(* IEC 61131-3 sources: brOscatLib/oscatBasic, 546 files *)

(* ---- oscatBasic.typ ---- *)
TYPE
    REAL2 :    STRUCT
        R1 : REAL; (* small value *)
        RX : REAL; (* big value *)
    END_STRUCT;
    CONSTANTS_LANGUAGE :    STRUCT
        DEFAULT : INT := 1; (* 1=english, 2=german 3=french *)
        LMAX : INT := 3;
        WEEKDAYS : ARRAY[1..3, 1..7] OF STRING[10] := ['Monday', 'Tuesday', 'Wednesday', 'Thursday', 'Friday', 'Saturday', 'Sunday', 'Montag', 'Dienstag', 'Mittwoch', 'Donnerstag', 'Freitag', 'Samstag', 'Sonntag', 'Lundi', 'Mardi', 'Mercredi', 'Jeudi', 'Vendredi', 'Samedi', 'Dimanche'];
        WEEKDAYS2 : ARRAY[1..3, 1..7] OF STRING[2] := ['Mo', 'Tu', 'We', 'Th', 'Fr', 'Sa', 'Su', 'Mo', 'Di', 'Mi', 'Do', 'Fr', 'Sa', 'So', 'Lu', 'Ma', 'Me', 'Je', 'Ve', 'Sa', 'Di'];
        MONTHS : ARRAY[1..3, 1..12] OF STRING[10] := ['January', 'February', 'March', 'April', 'May', 'June', 'July', 'August', 'September', 'October', 'November', 'December', 'Januar', 'Februar', 'März', 'April', 'Mai', 'Juni', 'Juli', 'August', 'September', 'Oktober', 'November', 'Dezember', 'Janvier', 'Février', 'mars', 'Avril', 'Mai', 'Juin', 'Juillet', 'Août', 'Septembre', 'Octobre', 'Novembre', 'Decembre'];
        MONTHS3 : ARRAY[1..3, 1..12] OF STRING[3] := ['Jan', 'Feb', 'Mar', 'Apr', 'May', 'Jun', 'Jul', 'Aug', 'Sep', 'Oct', 'Nov', 'Dec', 'Jan', 'Feb', 'Mrz', 'Apr', 'Mai', 'Jun', 'Jul', 'Aug', 'Sep', 'Okt', 'Nov', 'Dez', 'Jan', 'Fev', 'Mar', 'Avr', 'Mai', 'Jun', 'Jul', 'Aou', 'Sep', 'Oct', 'Nov', 'Dec'];
        DIRS : ARRAY[1..3, 0..15] OF STRING[3] := ['N', 'NNE', 'NE', 'ENE', 'E', 'ESE', 'SE', 'SSE', 'S', 'SSW', 'SW', 'WSW', 'W', 'WNW', 'NW', 'NNW', 'N', 'NNO', 'NO', 'ONO', 'O', 'OSO', 'SO', 'SSO', 'S', 'SSW', 'SW', 'WSW', 'W', 'WNW', 'NW', 'NNW', 'N', 'NNO', 'NO', 'ONO', 'O', 'OSO', 'SO', 'SSO', 'S', 'SSW', 'SW', 'WSW', 'W', 'WNW', 'NW', 'NNW'];
    END_STRUCT;
    CONSTANTS_LOCATION :    STRUCT
        DEFAULT : INT := 1; (* 1=germany, 2=austria 3=france 4=belgium-german 5= italien-Südtirol *)
        LMAX : INT := 5;
        LANGUAGE : ARRAY[1..5] OF INT := [2, 2, 3, 2, 2]; (* language spoken in the location *)
    END_STRUCT;
    CONSTANTS_MATH :    STRUCT
        PI : REAL := 3.1415926535897931; (* Kreiszahl PI *)
        PI2 : REAL := 6.2831853071795862; (* PI * 2 *)
        PI4 : REAL := 12.566370614359172; (* PI * 4 *)
        PI05 : REAL := 1.5707963267949; (* PI / 2 *)
        PI025 : REAL := 0.785398163397448; (* PI / 4 *)
        PI_INV : REAL := 0.318309886183791; (* 1 / PI *)
        E : REAL := 2.7182818284590451; (* Euler constant e *)
        E_INV : REAL := 0.367879441171442; (* 1 / e *)
        SQ2 : REAL := 1.4142135623731; (* Wurzel von 2 *)
        FACTS : ARRAY[0..12] OF DINT := [1, 1, 2, 6, 24, 120, 720, 5040, 40320, 362880, 3628800, 39916800, 479001600];
    END_STRUCT;
    CONSTANTS_PHYS :    STRUCT
        C : REAL := 299792458; (* Lichtgeschwindigkeit in m/s *)
        E : REAL := 1.60217653E-19; (* elementarladung in Colomb = A * s *)
        G : REAL := 9.80665; (* Erdbeschleunigung in m / s² *)
        T0 : REAL := -273.15; (* absoluter Nullpunkt in °C *)
        RU : REAL := 8.314472; (* Universelle Gaskonstante in J / (mol · K) *)
        PN : REAL := 101325; (* NormalDruck in Pa *)
    END_STRUCT;
    CONSTANTS_SETUP :    STRUCT
        EXTENDED_ASCII : BOOL := TRUE; (* setup Parameters *)
        CHARNAMES : ARRAY[1..4] OF STRING[253] := [';"&quot;&&amp;<&lt;>&gt;€&euro; &nbsp;¡&iexcl;¢&cent;£&pound;¤&curren;¥&yen;¦&brvbar;§&sect;¨&uml;©&copy;ª&ordf;«&laquo;¬&not;­&shy;®&reg;¯&macr;°&deg;±&plusmn;²&sup2;³&sup3;´&acute;µ&micro;¶&para;·&middot;¸&cedil;¹&sup1;º&ordm;»&raquo;¼&frac14;Û&Ucirc;',
		';¾&frac34;¿&iquest;À&Agrave;Á&Aacute;Â&Acirc;Ã&Atilde;Ä&Auml;Å&Aring;Æ&AElig;Ç&Ccedil;È&Egrave;É&Eacute;Ê&Ecirc;Ë&Euml;Ì&Igrave;Í&Iacute;Î&Icirc;Ï&Iuml;Ð&ETH;Ñ&Ntilde;Ò&Ograve;Ó&Oacute;Ô&Ocirc;Õ&Otilde;Ö&Ouml;×&times;Ø&Oslash;Ù&Ugrave;Ú&Uacute;½&frac12;',
		';Ü&Uuml;Ý&Yacute;Þ&THORN;ß&szlig;à&agrave;á&aacute;â&acirc;ã&atilde;ä&auml;å&aring;æ&aelig;ç&ccedil;è&egrave;é&eacute;ê&ecirc;ë&euml;ì&igrave;í&iacute;î&icirc;ï&iuml;ð&eth;ñ&ntilde;ò&ograve;ó&oacute;ô&ocirc;õ&otilde;ö&ouml;÷&divide;ø&oslash;ù&ugrave;',
		';ú&uacute;û&ucirc;ü&uuml;ý&yacute;þ&thorn;ÿ&yuml;'];
        MTH_OFS : ARRAY[1..12] OF INT := [0, 31, 59, 90, 120, 151, 181, 212, 243, 273, 304, 334];
        DECADES : ARRAY[0..8] OF REAL := [1, 10, 100, 1000, 10000, 100000, 1000000, 10000000, 100000000];
    END_STRUCT;
    TIMER_EVENT :    STRUCT
        TYP : BYTE;
        CHANNEL : BYTE;
        DAY : BYTE;
        START : TOD;
        DURATION : TIME;
        LAND : BYTE;
        LOR : BYTE;
        LAST : DT;
    END_STRUCT;
    FRACTION :    STRUCT
        NUMERATOR : INT;
        DENOMINATOR : INT;
    END_STRUCT;
    COMPLEX :    STRUCT
        re : REAL;
        im : REAL;
    END_STRUCT;
    VECTOR_3 :    STRUCT
        X : REAL;
        Y : REAL;
        Z : REAL;
    END_STRUCT;
    ESR_DATA :    STRUCT
        TYP : BYTE;
        ADRESS : STRING[10];
        DS : DT;
        TS : TIME;
        DATA : ARRAY[0..7] OF BYTE;
    END_STRUCT;
    CALENDAR :    STRUCT
        UTC : DT; (* world time UTC *)
        LOCAL_DT : DT; (* local time *)
        LOCAL_DATE : DATE; (* local date *)
        LOCAL_TOD : TOD; (* local time of day *)
        YEAR : INT; (* year of LDATE *)
        MONTH : INT; (* month of LDATE *)
        DAY : INT; (* day of LDATE *)
        WEEKDAY : INT; (* weekday of LDATE *)
        OFFSET : INT; (* Time Zone Offset for Local time in minutes *)
        DST_EN : BOOL; (* daylight savings time enable *)
        DST_ON : BOOL; (* true when daylight savings time os on *)
        NAME : STRING[5]; (* name of time zone *)
        LANGUAGE : INT; (* location number pls see location setup *)
        LONGITUDE : REAL; (* longitude of current location *)
        LATITUDE : REAL; (* latitude of current location *)
        SUN_RISE : TOD; (* sun_rise for current location *)
        SUN_SET : TOD; (* sun_set for current location *)
        SUN_MIDDAY : TOD; (* worldtime when sun stands at south position *)
        SUN_HEIGTH : REAL; (* suns heigth at midday, south position *)
        SUN_HOR : REAL; (* sun angle horizontal 0 = north in degrees *)
        SUN_VER : REAL; (* sun angle vertical above horizon in degrees *)
        NIGHT : BOOL; (* true between sun_set and sun_rise *)
        HOLIDAY : BOOL; (* true when holiday *)
        HOLY_NAME : STRING[30]; (* name of holiday *)
        WORK_WEEK : INT; (* current work week *)
    END_STRUCT;
    HOLIDAY_DATA :    STRUCT
        NAME : STRING[30];
        DAY : SINT;
        MONTH : SINT;
        USE : SINT;
    END_STRUCT;
    SDT :    STRUCT
        YEAR : INT;
        MONTH : INT;
        DAY : INT;
        WEEKDAY : INT;
        HOUR : INT;
        MINUTE : INT;
        SECOND : INT;
        MS : INT;
    END_STRUCT;
END_TYPE

(* ---- _ARRAY_ABS.st ---- *)
FUNCTION _ARRAY_ABS
    (*http://www.oscat.de/images/OSCATBasic/oscat_basic333_en.pdf#page=71*)
    stop := SHR(SIZE,2)-1;
    FOR i := 0 TO stop DO
    	PT[i] := ABS(PT[i]);
    END_FOR
    _ARRAY_ABS := TRUE;

    (* revision history
    hm	2. apr 2008		rev 1.0
    	original version

    *)
END_FUNCTION

(* ---- _ARRAY_ADD.st ---- *)
FUNCTION _ARRAY_ADD
    (*http://www.oscat.de/images/OSCATBasic/oscat_basic333_en.pdf#page=71*)
    stop := SHR(SIZE,2)-1;
    FOR i := 0 TO stop DO
    	PT[i] := PT[i] + X;
    END_FOR
    _ARRAY_ADD := TRUE;

    (* revision history
    hm	2. apr 2008		rev 1.0
    	original version

    *)
END_FUNCTION

(* ---- _ARRAY_INIT.st ---- *)
FUNCTION _ARRAY_INIT
    (*http://www.oscat.de/images/OSCATBasic/oscat_basic333_en.pdf#page=72*)
    stop := SHR(SIZE,2)-1;
    FOR i := 0 TO stop DO
    	PT[i] := INIT;
    END_FOR

    _ARRAY_INIT := TRUE;

    (* revision History

    hm 6.1.2007		rev 1.1
    	change type of function to bool
    	added  array_init := true to set output true.

    hm	14.11.2007	rev 1.2
    	changed stop calculation to be more efficient

    hm	16.3. 2008		rev 1.3
    	changed type of input SIZE to uint
    *)
END_FUNCTION

(* ---- _ARRAY_MEDIAN.st ---- *)
FUNCTION _ARRAY_MEDIAN
    (*http://www.oscat.de/images/OSCATBasic/oscat_basic333_en.pdf#page=73*)
    _ARRAY_SORT(ADR(PT),SIZE);
    stop := SHR(SIZE,2)-1;
    IF EVEN(UINT_TO_INT(stop)) THEN
    	_ARRAY_MEDIAN := PT[SHR(stop,1)];
    ELSE
    	i := SHR(stop,1);
    	_ARRAY_MEDIAN := (PT[i] + PT[i+1]) * 0.5;
    END_IF

    (* old code
    stop := (SIZE - SIZEOF(PT)) / SIZEOF(PT);
    FOR i := 0 TO stop - 1 DO
    	FOR m := i + 1 TO stop DO
    		IF PT[i] > PT[m] THEN
    			temp := PT[i];
    			PT[i] := PT[m];
    			PT[m] := temp;
    		END_IF
    	END_FOR
    END_FOR
    IF even(stop) THEN
    	_ARRAY_MEDIAN := PT[stop/2];
    ELSE
    	i := stop/2;
    	_ARRAY_MEDIAN := (PT[i] + PT[i+1])/2;
    END_IF
    *)
    (* revision history
    hm 	3.3.2007		rev 1.1
    	corrected an error, changed the statement line 14	i := TRUNC(stop/2); to i := stop/2;

    hm		22. sep 2007	rev 1.2
    	changed algorithm to use _array_soft for performance reasons

    hm		8. oct 2007		rev 1.3
    	deleted unused variables m and temp

    hm		14. nov 2007	rev 1.4
    	corrected a problem with SIZE calculation

    hm		16.3. 2008		rev 1.5
    	changed type of input SIZE to uint
    	performance improvements
    *)
END_FUNCTION

(* ---- _ARRAY_MUL.st ---- *)
FUNCTION _ARRAY_MUL
    (*http://www.oscat.de/images/OSCATBasic/oscat_basic333_en.pdf#page=73*)
    stop := SHR(SIZE,2)-1;
    FOR i := 0 TO stop DO
    	PT[i] := PT[i] * X;
    END_FOR
    _ARRAY_MUL := TRUE;

    (* revision history
    hm	2. apr 2008		rev 1.0
    	original version

    *)
END_FUNCTION

(* ---- _ARRAY_SHUFFLE.st ---- *)
FUNCTION _ARRAY_SHUFFLE
    (*http://www.oscat.de/images/OSCATBasic/oscat_basic333_en.pdf#page=74*)
    stop := UINT_TO_INT(SHR(SIZE,2)-1);
    FOR i := 0 TO stop DO
            pos := RDM2(i+pos,0,stop);
            (* swap elements *)
            temp := PT[i];
            PT[i] := PT[pos];
            PT[pos] := temp;
    END_FOR

    _ARRAY_SHUFFLE := TRUE;

    (* revision History
    hm 	4. mar 2008	rev 1.0
    	original version

    hm	16. mar. 2008	rev 1.1
    	changed type of input SIZE to uint

    hm	30. mar. 2008	rev 1.2
    	changed last in rdm2 fromm pos to i + pos to allow for more randomness

    *)
END_FUNCTION

(* ---- _ARRAY_SORT.st ---- *)
FUNCTION _ARRAY_SORT
    (*http://www.oscat.de/images/OSCATBasic/oscat_basic333_en.pdf#page=75*)
    (* Startwerte zur Arraygröße *)
    links := 1;					(* Anfangselement des Arrays *)
    rechts := SHR(SIZE,2);		(* Endelement des Arrays *)
    stack_count := 1;			(* Laufvariable stack *)

    WHILE NOT ende_aussen DO						(* äußere Schleife *)
    	IF links < rechts THEN
    		pivot := PT[SHR(rechts+links,1)];			(* Wert des mittleren Elements als pivot-Wert *)
    		i := links -1;
    		j := rechts +1;

    		(* innere Schleife, teile Feld *)
    		ende_innen := FALSE;
    		REPEAT

    			(* steigende Reihenfolge *)
    			REPEAT	i := i+1;	UNTIL (PT[i] >= pivot) OR NOT (i < rechts)	END_REPEAT
    			REPEAT	j := j-1;	UNTIL (PT[j] <= pivot) OR NOT (j > links)	END_REPEAT

    			(*sinkende Reihenfolge *)
    (*			REPEAT	i := i+1;	UNTIL (PT[i] <= pivot) OR NOT (i < rechts)	END_REPEAT	*)
    (*			REPEAT	j := j-1;	UNTIL (PT[j] >= pivot) OR NOT (j > links)	END_REPEAT	*)

    			IF i >= j THEN
    				ende_innen := TRUE;
    			ELSE
    				   tmp := PT[j];
    				PT[j] := PT[i];
    				PT[i] := tmp;
    			END_IF

    		UNTIL ende_innen END_REPEAT

    		(* Push stack *)
    		stack[stack_count] := rechts;		(* rechten Teil später sortieren *)
    		IF stack_count < 32 THEN
    			stack_count := stack_count +1;
    		ELSE
    			ende_aussen := TRUE;
    			_ARRAY_SORT := FALSE;					(* Fehler: stack zu klein *)
    		END_IF

    		(* linken Teil sortiern *)
    		rechts := MAX(links, i-1);

    	ELSE

    		IF stack_count = 1 THEN
    			ende_aussen := TRUE;
    		ELSE

    			links := rechts+1;

    			(* pop stack *)
    			stack_count := stack_count -1;		(* jetzt rechten Teil sortierne *)
    			rechts:= stack[stack_count];
    		END_IF

    	END_IF

    END_WHILE

    _ARRAY_SORT := TRUE;				(* Sortierung beendet *)

    (* algorithm used before rev 2.0

    SIZE := SHR(SIZE,2);
    size2 := UINT_TO_INT(SHR(SIZE,1));
    FOR i := SIZE2  TO 1 BY -1 DO
    	j:=i;
        WHILE j <= SIZE2 DO
         	stop := j * 2 + 1;
            IF stop > UINT_TO_INT(SIZE) THEN stop := stop - 1;
            ELSIF PT[stop-1] > PT[stop] THEN stop := stop - 1;
    		END_IF
            IF PT[j] < PT[stop] THEN
             	temp := PT[j];
                PT[j] := PT[stop];
                PT[stop] := temp;
            END_IF
            j := stop;
        END_WHILE
    END_FOR

    *)

    (* heapsort
    FOR heapsize := UINT_TO_INT(SIZE) TO 1 BY -1 DO
    	popmax := PT[1];
    	PT[1] := PT[heapsize];
       	i := 1;
    	hs2 := SHR(heapsize,1);
    	WHILE i <= hs2 DO
           	stop := i * 2 + 1;
            	IF stop > heapsize THEN stop := stop - 1;
            	ELSIF PT[stop-1] > PT[stop] THEN stop := stop - 1;
    	 	END_IF
            	IF PT[i] < PT[stop] THEN
                		temp := PT[i];
                		PT[i] := PT[stop];
                		PT[stop] := temp;
            	END_IF
            	i := stop;
        	END_WHILE
    	PT[heapsize] := popmax;
    END_FOR

    _ARRAY_SORT2 := TRUE;
    *)

    (* old algorithm bubble sort used before rev 1.2
    stop := (SIZE - SIZEOF(PT)) / SIZEOF(PT);
    FOR i := 0 TO stop - 1 DO
    	FOR m := i + 1 TO stop DO
    		IF PT[i] > PT[m] THEN
    			temp := PT[i];
    			PT[i] := PT[m];
    			PT[m] := temp;
    		END_IF
    	END_FOR
    END_FOR
    _ARRAY_SORT := TRUE;

    *)

    (* revision history

    hm 	6.1.2007 	rev 1.1
    	changed return value to true

    hm	22. sep 2007	rev 1.2
    	changed sorting algorithm to heap sort for performance reasons

    hm 	14. nov 2007	rev 1.3
    	changed calculation of stop to be more efficient

    hm	15 dec 2007	rev 1.4
    	added function return true

    hm	5. jan 2008		rev 1.5
    	improved performance

    hm	16. mar. 2008	rev 1.6
    	changed type of input SIZE to uint

    hm	28. mar. 2008	rev 1.7
    	changed input f to PT

    hm	19. jan. 2011	rev 2.0
    	new faster algorithm using qucksort (Alexander Drikitis)

    *)

END_FUNCTION

(* ---- _BUFFER_CLEAR.st ---- *)
FUNCTION _BUFFER_CLEAR
    (*http://www.oscat.de/images/OSCATBasic/oscat_basic333_en.pdf#page=477*)
    (* this routine uses 32 bit access to gain speed *)
    (* first access bytes till pointer is aligned for 32 bit access *)
    temp := ADR(PT);
    end := temp + SIZE;
    end32 := end - 3;
    WHILE (ADR(PT) < end) AND ((temp AND 16#00000003) > 0) DO
    	PT := 0;
    	PT ACCESS (ADR(PT) + 1);
    	temp := temp + 1;
    END_WHILE
    (* pointer is aligned, now copy 32 bits at a time *)
    ptw ACCESS ADR(PT);
    WHILE ADR(ptw) < end32 DO (* *)
    	ptw := 0;
    	ptw ACCESS (ADR(ptw) + 4);
    END_WHILE
    (* copy the remaining bytes in byte mode *)
    PT ACCESS ADR(ptw);
    WHILE ADR(PT) < end DO
    	PT := 0;
    	PT ACCESS (ADR(PT) + 1);
    END_WHILE

    _BUFFER_CLEAR := TRUE;

    (* revision History
    hm 	5. mar. 2008	rev 1.0
    	original version

    hm	16. mar. 2008	rev 1.1
    	added type conversion to avoid warnings under codesys 30
    	chaged type of input SIZE to uint
    	deleted unused variable i

    hm	31. oct. 2008	rev 1.2
    	corrected an error while routine would write outside of arrays

    *)
END_FUNCTION

(* ---- _BUFFER_INIT.st ---- *)
FUNCTION _BUFFER_INIT
    (*http://www.oscat.de/images/OSCATBasic/oscat_basic333_en.pdf#page=477*)
    (* this routine uses 32 bit access to gain speed *)
    (* first access bytes till pointer is aligned for 32 bit access *)
    temp := ADR(PT);
    end := temp + SIZE;
    end32 := end - 3;
    WHILE (ADR(PT) < end) AND ((temp AND 16#00000003) > 0) DO
    	PT := INIT;
        PT ACCESS (ADR(PT) + 1);
    	temp := temp + 1;
    END_WHILE
    (* pointer is aligned, now copy 32 bits at a time *)
    ptw ACCESS ADR(PT);
    temp := SHL(BYTE_TO_UDINT(INIT),24) OR SHL(BYTE_TO_UDINT(INIT),16) OR SHL(BYTE_TO_UDINT(INIT),8) OR BYTE_TO_UDINT(INIT);
    WHILE ADR(ptw) < end32 DO
    	ptw := UDINT_TO_DWORD(temp);
    	ptw ACCESS (ADR(ptw) + 4);
    END_WHILE
    (* copy the remaining bytes in byte mode *)
    PT ACCESS ADR(ptw);
    WHILE ADR(PT) < end DO
    	PT := INIT;
    	PT ACCESS (ADR(PT) + 1);
    END_WHILE

    _BUFFER_INIT := TRUE;

    (* revision History
    hm 	5. mar. 2008	rev 1.0
    	original version

    hm	16. mar. 2008	rev 1.1
    	added type conversion to avoid warnings under codesys 3.0
    	chaged type of input SIZE to uint.

    hm	31. oct. 2008	rev 1.2
    	corrected an error while routine would write outside of arrays

    *)
END_FUNCTION

(* ---- _BUFFER_INSERT.st ---- *)
FUNCTION _BUFFER_INSERT
    (*http://www.oscat.de/images/OSCATBasic/oscat_basic333_en.pdf#page=478*)
    lx := LEN(STR);
    end := POS + lx;
    (* first move the upper part of the buffer to make space for the string *)
    FOR i := UINT_TO_INT(SIZE) - 1 TO end BY -1 DO
    	PT[i] := PT[i-lx];
    END_FOR
    (* copy the string *)
    _BUFFER_INSERT := _STRING_TO_BUFFER(STR, POS, ADR(PT), SIZE);

    (* revision History
    hm 	9. mar. 2008	rev 1.0
    	original version

    hm	16. mar. 2008	rev 1.1
    	changed type of input SIZE to uint

    hm	13. may. 2008	rev 1.2
    	changed type of pointer to array[1..32767]
    	changed SIZE of string to STRING_LENGTH

    hm	23. mar. 2009	rev 1.3
    	avoid writing to input POS

    hm	12. nov. 2009	rev 1.4
    	code optimized

    hm 2. jan 2012	rev 1.5
    	function now returns the next position after the input string

    *)
END_FUNCTION

(* ---- _BUFFER_UPPERCASE.st ---- *)
FUNCTION _BUFFER_UPPERCASE
    (*http://www.oscat.de/images/OSCATBasic/oscat_basic333_en.pdf#page=479*)
    pos := 0;
    WHILE pos < SIZE DO
    	PT[pos] := TO_UPPER(PT[pos]);
    	pos := pos + 1;
    END_WHILE

    _BUFFER_UPPERCASE := TRUE;

    (* revision History
    hm 	20. jan. 2011	rev 1.0
    	original version

    *)
END_FUNCTION

(* ---- _STRING_TO_BUFFER.st ---- *)
FUNCTION _STRING_TO_BUFFER
    (*http://www.oscat.de/images/OSCATBasic/oscat_basic333_en.pdf#page=479*)
    ps ACCESS ADR(STR);
    end := MIN(POS + LEN(STR), UINT_TO_INT(SIZE));
    IF end > 0 THEN end := end -1; END_IF
    FOR i := POS TO end DO
    	PT[i] := ps;
    	ps ACCESS (ADR(ps) + 1);
    END_FOR

    _STRING_TO_BUFFER := i;

    (* revision History

    hm 	5. mar. 2008	rev 1.0
    	original version

    hm	16. mar. 2008	rev 1.1
    	changed type of input SIZE to uint

    hm	13. may. 2008	rev 1.2
    	changed type of pointer to array[1..32767]
    	changed SIZE of string to STRING_LENGTH

    hm	12. nov. 2009	rev 1.3
    	limit end to SIZE - 1

    hm	2. jan 2012	rev 1.4
    	return the position after the input string when finished
    *)
END_FUNCTION

(* ---- ACOSH.st ---- *)
FUNCTION ACOSH
    (*http://www.oscat.de/images/OSCATBasic/oscat_basic333_en.pdf#page=39*)
    ACOSH := LN(SQRT(X * X - 1.0) + X);

    (* revision history
    hm		12 jan 2007	rev 1.0
    	original version

    hm		2. dec 2007	rev 1.1
    	changed code for better performance

    hm	16. mar. 2007		rev 1.2
    	changed sequence of calculations to improve performance

    hm	10. mar. 2009		rev 1.3
    	real constants updated to new systax using dot

    *)
END_FUNCTION

(* ---- ACOTH.st ---- *)
FUNCTION ACOTH
    (*http://www.oscat.de/images/OSCATBasic/oscat_basic333_en.pdf#page=39*)
    ACOTH := LN((X+1.0)/(X-1.0))*0.5;

    (* revision history
    hm		12 jan 2007	rev 1.0
    	original version

    hm		5. jan 2008	rev 1.1
    	improved code for better performance

    hm	10. mar. 2009		rev 1.2
    	real constants updated to new systax using dot

    *)
END_FUNCTION

(* ---- AGDF.st ---- *)
FUNCTION AGDF
    (*http://www.oscat.de/images/OSCATBasic/oscat_basic333_en.pdf#page=39*)
    AGDF := LN((1.0 + SIN(X)) / COS(X));

    (* comment
    the current implementation gives sufficient accuracy only up to X = 1.57 or an output > 10.
    is X closer to PI/2 then the function is more and more unreliable
    *)

    (* revision history
    hm	27. apr. 2008	rev 1.0
    	original version

    hm	10. mar. 2009	rev 1.1
    	real constants updated to new systax using dot

    *)

END_FUNCTION

(* ---- AIN.st ---- *)
FUNCTION AIN
    (*http://www.oscat.de/images/OSCATBasic/oscat_basic333_en.pdf#page=269*)
    (* extract the SIGN bit *)
    IF SIGN < 32 THEN
    	temp1 := SHR(IN,SIGN);
    	sx := temp1.0;
    ELSE
    	sx := FALSE;
    END_IF
    temp1 := SHR(ff, 32-BYTE_TO_USINT(BITS));
    temp2 := IN AND temp1;
    AIN := (HIGH - LOW) * DWORD_TO_REAL(temp2) / DWORD_TO_REAL(temp1) + LOW;
    IF sx THEN AIN := -AIN; END_IF

    (* revision history
    hm 18.8.2006	rev 1.1
    	fixed an error with LOW value negative and HIGH value 0.

    hm 19.1.2007	rev 1.2
    	fixed an error with SIGN bit.

    hm	13.9.2007	rev 1.3
    	changed code to avoid warning under codesys 2.8.1

    hm	2. dec 2007	rev 1.4
    	changed code for better performance

    hm	16. mar 2008	rev 1.5
    	added type conversions to avoid warnings under codesys 30
    *)
END_FUNCTION

(* ---- AOUT.st ---- *)
FUNCTION AOUT
    (*http://www.oscat.de/images/OSCATBasic/oscat_basic333_en.pdf#page=271*)
    (* if SIGN bit is defined *)
    IF SIGN < 32 THEN
    	sx := SIGN_R(IN);
    	in2 := ABS(IN);
    ELSE
    	in2 := IN;
    END_IF

    (* begrenze IN auf die zulässigen werte *)
    in2 := LIMIT(LOW, in2, HIGH);

    (* Berechne den Ausgangswert *)
    AOUT := REAL_TO_DWORD((in2 - LOW) / (HIGH - LOW) * UDINT_TO_REAL(SHL(ff,BYTE_TO_USINT(BITS)) -1));
    IF sx THEN AOUT := UDINT_TO_DWORD(SHL(ff,SIGN) OR DWORD_TO_UDINT(AOUT)); END_IF

    (*
    revision history

    hm 18.1.2007		rev 1.1
    	renamed Modul to AOUT.
    	changed Output to 32 Bit max.
    	corrected error with SIGN bit.

    hm	13.9.2007		rev 1.2
    	changed code to avoid warning under codesys 2.8.1

    hm	2. dec 2007		rev 1.3
    	changed code for better performance

    hm	23. feb 2008	rev 1.4
    	changed code for better performance
    *)
END_FUNCTION

(* ---- AOUT1.st ---- *)
FUNCTION AOUT1
    (*http://www.oscat.de/images/OSCATBasic/oscat_basic333_en.pdf#page=272*)
    (* if SIGN bit is defined *)
    IF SIGN < 32 THEN
    	sx := SIGN_R(IN);
    	in2 := ABS(IN);
    ELSE
    	in2 := IN;
    END_IF

    (* begrenze IN auf die zulässigen werte *)
    in2 := LIMIT(LOW, in2, HIGH);

    (* Berechne den Ausgangswert *)
    AOUT1 := SHL(REAL_TO_DWORD((in2 - LOW) / (HIGH - LOW) * UDINT_TO_REAL(SHL(ff,BIT_N - BIT_0 + 1) -1)),BIT_0);
    IF sx THEN AOUT1 := UDINT_TO_DWORD(SHL(ff,SIGN) OR DWORD_TO_UDINT(AOUT1)); END_IF

    (* revision history
    hm	23. feb 2008	rev 1.0
    	original version

    *)
END_FUNCTION

(* ---- ARRAY_AVG.st ---- *)
FUNCTION ARRAY_AVG
    (*http://www.oscat.de/images/OSCATBasic/oscat_basic333_en.pdf#page=76*)
    stop := SHR(SIZE,2)-1;
    ARRAY_AVG := PT[0];
    FOR i := 1 TO stop DO
    	ARRAY_AVG := ARRAY_AVG + PT[i];
    END_FOR
    ARRAY_AVG := ARRAY_AVG / UINT_TO_REAL(stop + 1);

    (* revision history
    hm	2. oct 2007		rev 1.0
    	original version

    hm	12. dec 2007	rev 1.1
    	chaged code for better performance

    hm	16. mar. 2008	rev 1.2
    	changed input SIZE to uint

    hm	10. mar. 2009	rev 1.3
    	added type conversion for compatibility reasons
    *)
END_FUNCTION

(* ---- ARRAY_GAV.st ---- *)
FUNCTION ARRAY_GAV
    (*http://www.oscat.de/images/OSCATBasic/oscat_basic333_en.pdf#page=76*)
    stop := SHR(SIZE,2)-1;
    ARRAY_GAV := 1.0;
    FOR i := 0 TO stop DO
    	IF PT[i] > 0.0 THEN
    		ARRAY_GAV := ARRAY_GAV * PT[i];
    	ELSE
    		ARRAY_GAV := 0.0;
    		RETURN;
    	END_IF
    END_FOR
    ARRAY_GAV := SQRTN(ARRAY_GAV,UINT_TO_INT(stop)+1);

    (* revision history
    hm	2. apr 2008	rev 1.0
    	original version

    hm	10. mar. 2009	rev 1.1
    	real constants updated to new systax using dot

    *)
END_FUNCTION

(* ---- ARRAY_HAV.st ---- *)
FUNCTION ARRAY_HAV
    (*http://www.oscat.de/images/OSCATBasic/oscat_basic333_en.pdf#page=77*)
    stop := SHR(SIZE,2)-1;
    FOR i := 0 TO stop DO
    	IF PT[i] <> 0.0 THEN
    		ARRAY_HAV := ARRAY_HAV + 1.0 / PT[i];
    	ELSE
    		ARRAY_HAV := 0.0;
    		RETURN;
    	END_IF
    END_FOR
    ARRAY_HAV := UINT_TO_REAL(stop + 1) / ARRAY_HAV;

    (* revision history
    hm	2. apr 2008	rev 1.0
    	original version

    hm	10. mar. 2009	rev 1.1
    	real constants updated to new systax using dot

    *)
END_FUNCTION

(* ---- ARRAY_MAX.st ---- *)
FUNCTION ARRAY_MAX
    (*http://www.oscat.de/images/OSCATBasic/oscat_basic333_en.pdf#page=77*)
    stop := (SIZE -SIZEOF(PT)) / SIZEOF(PT);
    ARRAY_MAX := PT[0];
    FOR i := 1 TO stop DO
    	IF PT[i] > ARRAY_MAX THEN ARRAY_MAX := PT[i]; END_IF
    END_FOR

    (* revision history
    hm	2. oct 2006		rev 1.0
    	original version

    hm	16. mar. 2008	rev 1.1
    	changed input SIZE to uint
    *)
END_FUNCTION

(* ---- ARRAY_MIN.st ---- *)
FUNCTION ARRAY_MIN
    (*http://www.oscat.de/images/OSCATBasic/oscat_basic333_en.pdf#page=78*)
    stop := (SIZE - SIZEOF(PT)) / SIZEOF(PT);
    ARRAY_MIN := PT[0];
    FOR i := 1 TO stop DO
    	IF PT[i] < ARRAY_MIN THEN ARRAY_MIN := PT[i]; END_IF
    END_FOR

    (* revision history
    hm		2. oct. 2006
    	original version

    hm		16. mar. 2008
    	changed type of input SIZE to uint

    *)
END_FUNCTION

(* ---- ARRAY_SDV.st ---- *)
FUNCTION ARRAY_SDV
    (*http://www.oscat.de/images/OSCATBasic/oscat_basic333_en.pdf#page=79*)
    (* standard deviation is simply the square root of the variance *)

    ARRAY_SDV := SQRT(ARRAY_VAR(ADR(PT), SIZE));

    (* revision history
    hm 	1.4.2007		rev 1.0
    	function created

    hm	16. mar. 2008	rev 1.1
    	changed type of input SIZE to uint

    *)
END_FUNCTION

(* ---- ARRAY_SPR.st ---- *)
FUNCTION ARRAY_SPR
    (*http://www.oscat.de/images/OSCATBasic/oscat_basic333_en.pdf#page=79*)
    stop := (SIZE -SIZEOF(PT)) / SIZEOF(PT);
    array_min := PT[0];
    array_max := PT[0];
    FOR i := 1 TO stop DO
    	IF PT[i] > array_max THEN array_max := PT[i];
    	ELSIF PT[i] < array_min THEN array_min := PT[i];
    	END_IF
    END_FOR
    ARRAY_SPR := array_max - array_min;

    (* revision history
    hm 	2. oct. 2006	rev 1.0
    	original version

    hm	16. mar. 2008	rev 1.1
    	changed type of input SIZE to uint

    *)
END_FUNCTION

(* ---- ARRAY_SUM.st ---- *)
FUNCTION ARRAY_SUM
    (*http://www.oscat.de/images/OSCATBasic/oscat_basic333_en.pdf#page=80*)
    stop := (SIZE -SIZEOF(PT)) / SIZEOF(PT);
    ARRAY_SUM := PT[0];
    FOR i := 1 TO stop DO
    	ARRAY_SUM := ARRAY_SUM + PT[i];
    END_FOR

    (* revision history
    hm 	2. oct. 2006	rev 1.0
    	function created

    hm	16. mar. 2008	rev 1.1
    	changed type of input SIZE to uint

    *)
END_FUNCTION

(* ---- ARRAY_TREND.st ---- *)
FUNCTION ARRAY_TREND
    (*http://www.oscat.de/images/OSCATBasic/oscat_basic333_en.pdf#page=81*)
    stop := SHR(SIZE,2)-1;
    stop2 := SHR(stop,1);
    FOR i := 0 TO stop2 DO x := x - PT[i]; END_FOR
    IF EVEN(UINT_TO_INT(stop)) THEN
    	FOR i := stop2 TO stop DO x := x + PT[i]; END_FOR
    ELSE
    	FOR i := stop2 + 1 TO stop DO x := x + PT[i]; END_FOR
    END_IF
    ARRAY_TREND := x / UINT_TO_REAL(stop2 + 1);

    (* revision history
    hm	2 oct 2007	rev 1.0
    	original version

    hm	12 dec 2007	rev 1.1
    	changed code for better performance

    hm	16. mar. 2008	rev 1.2
    	changed type of input SIZE to uint

    hm	10. mar. 2009	rev 1.3
    	added type conversions for compatibility reasons
    *)
END_FUNCTION

(* ---- ARRAY_VAR.st ---- *)
FUNCTION ARRAY_VAR
    (*http://www.oscat.de/images/OSCATBasic/oscat_basic333_en.pdf#page=81*)
    (* at first we calualte the arithmetic average of the array *)

    stop := SHR(SIZE,2)-1;
    avg := PT[0];
    FOR i := 1 TO stop DO
    	avg := avg + PT[i];
    END_FOR
    avg := avg / UINT_TO_REAL(stop + 1);

    (* in a second run we calculate the variance of the array *)

    ARRAY_VAR := (PT[0] - avg) * (PT[0] - avg);
    FOR i := 1 TO stop DO
    	ARRAY_VAR := ARRAY_VAR + (PT[i] - avg) * (PT[i] - avg);
    END_FOR
    ARRAY_VAR := ARRAY_VAR / UINT_TO_REAL(stop);

    (* revision history
    hm 	1.4.2007	rev 1.0
    	function created

    hm	12.12.2007	rev 1.1
    	changed code for better performance

    hm	16. mar. 2008	rev 1.2
    	changed type of input SIZE to uint

    hm	10. mar. 2009	rev 1.3
    	added type conversions for compatibility reasons
    *)
END_FUNCTION

(* ---- ASINH.st ---- *)
FUNCTION ASINH
    (*http://www.oscat.de/images/OSCATBasic/oscat_basic333_en.pdf#page=40*)
    ASINH := LN(SQRT(X * X + 1.0)+X);

    (* revision history
    hm		12 jan 2007	rev 1.0
    	original version

    hm		2. dec 2007	rev 1.1
    	changed code for better performance

    hm		16.3. 2007		rev 1.2
    	changed sequence of calculations to improve performance

    hm	10. mar. 2009		rev 1.3
    	real constants updated to new systax using dot

    *)
END_FUNCTION

(* ---- ATAN2.st ---- *)
FUNCTION ATAN2
    (*http://www.oscat.de/images/OSCATBasic/oscat_basic333_en.pdf#page=40*)
    IF X > 0.0 THEN
    	ATAN2 := ATAN(Y/X);
    ELSIF X < 0.0 THEN
    	IF Y >=0.0 THEN
    		ATAN2 := ATAN(Y/X) + cPI;
    	ELSE
    		ATAN2 := ATAN(Y/X) - cPI;
    	END_IF
    ELSIF Y > 0.0 THEN
    	ATAN2 := cPI05;
    ELSIF Y < 0.0 THEN
    	ATAN2 := -cPI05;
    ELSE
    	ATAN2 := 0.0;
    END_IF

    (* revision history
    hm	20.  apr. 2008	rev 1.0
    	original version

    hm	18. oct. 2008	rev 1.1
    	changed to use math constants

    hm	10. mar. 2009	rev 1.2
    	real constants updated to new systax using dot

    *)

END_FUNCTION

(* ---- ATANH.st ---- *)
FUNCTION ATANH
    (*http://www.oscat.de/images/OSCATBasic/oscat_basic333_en.pdf#page=41*)
    ATANH := LN((1.0 + X)/(1.0 - X)) * 0.5;

    (* revision history
    hm		12 jan 2007	rev 1.0
    	original version

    hm		5. jan 2008	rev 1.1
    	improved code for better performance

    hm	10. mar. 2009		rev 1.2
    	real constants updated to new systax using dot

    *)

END_FUNCTION

(* ---- BAND_B.st ---- *)
FUNCTION BAND_B
    (*http://www.oscat.de/images/OSCATBasic/oscat_basic333_en.pdf#page=377*)
    IF BYTE_TO_SINT(X) < BYTE_TO_SINT(B) THEN
    	BAND_B := 0;
    ELSIF BYTE_TO_SINT(X) > (255 - BYTE_TO_SINT(B)) THEN
    	BAND_B := 255;
    ELSE
    	BAND_B := X;
    END_IF

    (* revision history
    hm	21. nov. 2008	rev 1.0
    	original version

    *)

END_FUNCTION

(* ---- BCDC_TO_INT.st ---- *)
FUNCTION BCDC_TO_INT
    (*http://www.oscat.de/images/OSCATBasic/oscat_basic333_en.pdf#page=210*)
    BCDC_TO_INT := (BYTE_TO_INT(IN) AND 16#0F) + (SHR(BYTE_TO_INT(IN),4) * 10);

    (* revision history
    hm	13.12.2007	rev 1.0
    	original version

    hm	30.6.2008	rev 1.1
    	changed name BCD_TO_INT to BCDC_TO_INT to avoid collision with util.lib

    *)
END_FUNCTION

(* ---- BETA.st ---- *)
FUNCTION BETA
    (*http://www.oscat.de/images/OSCATBasic/oscat_basic333_en.pdf#page=41*)
    BETA := GAMMA(X) * GAMMA(Y) / GAMMA(X + Y);

    (* revision history
    hm	26. oct. 2008	rev 1.0
    	original version

    *)
END_FUNCTION

(* ---- BFT_TO_MS.st ---- *)
FUNCTION BFT_TO_MS
    (*http://www.oscat.de/images/OSCATBasic/oscat_basic333_en.pdf#page=354*)
    BFT_TO_MS := EXPT(BFT, 1.5) * 0.836;

    (* revision history
    hm	12. 6. 2008		rev 1.0
    	original version

    *)
END_FUNCTION

(* ---- BIN_TO_BYTE.st ---- *)
FUNCTION BIN_TO_BYTE
    (*http://www.oscat.de/images/OSCATBasic/oscat_basic333_en.pdf#page=145*)
    pt ACCESS ADR(BIN);
    stop := LEN(BIN);
    FOR i := 1 TO stop DO
    	X := pt;
    	(* calculate the value of the digit *)
    	IF X = BYTE#48 THEN
    		BIN_TO_BYTE := SHL(BIN_TO_BYTE,1);
    	ELSIF X = BYTE#49 THEN
    		BIN_TO_BYTE := SHL(BIN_TO_BYTE,1) OR 1;
    	END_IF
    	pt ACCESS (ADR(pt) + 1);
    END_FOR

    (* revision histroy
    hm	18. jun. 2008	rev 1.0
    	original release

    hm	20. sep. 2008	rev 1.1
    	changed length of input string from 20 to 12

    hm	26. jul. 2009	rev 1.2
    	optimized code
    *)

END_FUNCTION

(* ---- BIN_TO_DWORD.st ---- *)
FUNCTION BIN_TO_DWORD
    (*http://www.oscat.de/images/OSCATBasic/oscat_basic333_en.pdf#page=145*)
    pt ACCESS ADR(BIN);
    stop := LEN(BIN);
    FOR i := 1 TO stop DO
    	X := pt;
    	(* calculate the value of the digit *)
    	IF X = BYTE#48 THEN
    		BIN_TO_DWORD := SHL(BIN_TO_DWORD,1);
    	ELSIF X = BYTE#49 THEN
    		BIN_TO_DWORD := SHL(BIN_TO_DWORD,1) OR 1;
    	END_IF
    	pt ACCESS (ADR(pt) + 1);
    END_FOR

    (* revision histroy
    hm	18. jun. 2008	rev 1.0
    	original release

    hm	20. sep. 2008	rev 1.1
    	changed length of input dtring from 20 to 40

    hm	26. jul 2009	rev 1.2
    	optimized code
    *)

END_FUNCTION

(* ---- BINOM.st ---- *)
FUNCTION BINOM
    (*http://www.oscat.de/images/OSCATBasic/oscat_basic333_en.pdf#page=42*)
    IF 2 * K > N THEN
    	K := N - K;
    END_IF
    IF K > N THEN
    	RETURN;
    ELSIF K = 0 OR K = N THEN
    	BINOM := 1;
    ELSIF K = 1 THEN
    	BINOM := N;
    ELSE
    	BINOM := N;
    	N := N + 1;
    	FOR i := 2 TO K DO
    		BINOM := BINOM * (N - i) / i;
    	END_FOR
    END_IF

    (*
    binomialkoeffizient(N, K)
    1  wenn K = 0 return 1
    2  wenn 2k > N
    3      dann führe aus ergebnis \leftarrow binomialkoeffizient(N, N-K)
    4  sonst führe aus ergebnis \leftarrow N
    5          von i \leftarrow 2 bis K
    6              führe aus ergebnis \leftarrow ergebnis \cdot (N + 1 - i)
    7                        ergebnis \leftarrow ergebnis : i
    8  return ergebnis
    *)

    (* revision history
    hm	25. oct. 2008	rev 1.0
    	original version

    *)
END_FUNCTION

(* ---- BIT_COUNT.st ---- *)
FUNCTION BIT_COUNT
    (*http://www.oscat.de/images/OSCATBasic/oscat_basic333_en.pdf#page=210*)
    WHILE IN > 0 DO
    	IF IN.0 THEN BIT_COUNT := BIT_COUNT + 1; END_IF
    	IN := SHR(IN,1);
    END_WHILE

    (* revision history
    5.7.2007	rev 1.0		original version

    10.9.2007	rev 1.1		hm
    	changed algorithm for better performace
    	the execution time has reduced by a factor of 5
    	deleted unused variable temp
    *)
END_FUNCTION

(* ---- BIT_LOAD_B.st ---- *)
FUNCTION BIT_LOAD_B
    (*http://www.oscat.de/images/OSCATBasic/oscat_basic333_en.pdf#page=210*)
    IF VAL THEN
    	BIT_LOAD_B := IN OR SHL(dat,POS);
    ELSE
    	BIT_LOAD_B := IN AND (NOT SHL(dat,POS));
    END_IF

    (* revision history
    hm	29. feb 2008	rev 1.0
    	original version

    hm	16. mar 2008	rev 1.1
    	change input bit to VAL for compatibility reasons
    *)

END_FUNCTION

(* ---- BIT_LOAD_B2.st ---- *)
FUNCTION BIT_LOAD_B2
    (*http://www.oscat.de/images/OSCATBasic/oscat_basic333_en.pdf#page=211*)
    IF D THEN
    	BIT_LOAD_B2 := ROL(SHR(BYTE#255, 8 - N) OR ROR(I, P), P);
    ELSE
    	BIT_LOAD_B2 := ROL(SHL(BYTE#255, N) AND ROR(I, P), P);
    END_IF

    (* revision history
    hm	18. oct. 2008	rev 1.0
    	original version

    *)

END_FUNCTION

(* ---- BIT_LOAD_DW.st ---- *)
FUNCTION BIT_LOAD_DW
    (*http://www.oscat.de/images/OSCATBasic/oscat_basic333_en.pdf#page=211*)
    IF VAL THEN
    	BIT_LOAD_DW := IN OR SHL(dat,POS);
    ELSE
    	BIT_LOAD_DW := IN AND (NOT SHL(dat,POS));
    END_IF

    (* revision history
    hm	29. feb 2008	rev 1.0
    	original version

    hm	16. mar 2008	rev 1.1
    	change input bit to VAL for compatibility reasons
    *)

END_FUNCTION

(* ---- BIT_LOAD_DW2.st ---- *)
FUNCTION BIT_LOAD_DW2
    (*http://www.oscat.de/images/OSCATBasic/oscat_basic333_en.pdf#page=212*)
    IF D THEN
    	BIT_LOAD_DW2 := ROL(SHR(DWORD#4294967295, 32 - N) OR ROR(I, P), P);
    ELSE
    	BIT_LOAD_DW2 := ROL(SHL(DWORD#4294967295, N) AND ROR(I, P), P);
    END_IF

    (* revision history
    hm	18. oct. 2008	rev 1.0
    	original version

    *)

END_FUNCTION

(* ---- BIT_LOAD_W.st ---- *)
FUNCTION BIT_LOAD_W
    (*http://www.oscat.de/images/OSCATBasic/oscat_basic333_en.pdf#page=212*)
    IF VAL THEN
    	BIT_LOAD_W := IN OR SHL(dat,POS);
    ELSE
    	BIT_LOAD_W := IN AND (NOT SHL(dat,POS));
    END_IF

    (* revision history
    hm	29. feb 2008	rev 1.0
    	original version

    hm	16. mar 2008	rev 1.1
    	change input bit to VAL for compatibility reasons
    *)

END_FUNCTION

(* ---- BIT_LOAD_W2.st ---- *)
FUNCTION BIT_LOAD_W2
    (*http://www.oscat.de/images/OSCATBasic/oscat_basic333_en.pdf#page=213*)
    IF D THEN
    	BIT_LOAD_W2 := ROL(SHR(WORD#65535, 16 - N) OR ROR(I, P), P);
    ELSE
    	BIT_LOAD_W2 := ROL(SHL(WORD#65535, N) AND ROR(I, P), P);
    END_IF

    (* revision history
    hm	18. oct. 2008	rev 1.0
    	original version

    *)

END_FUNCTION

(* ---- BIT_OF_DWORD.st ---- *)
FUNCTION BIT_OF_DWORD
    (*http://www.oscat.de/images/OSCATBasic/oscat_basic333_en.pdf#page=213*)
    BIT_OF_DWORD := (SHR(IN,N) AND 16#00000001) > 0;

    (* old code used before rev 1.1
    temp := SHR(IN,N);
    BIT_OF_DWORD := temp.0;
    *)

    (* revision history
    hm	4. aug. 2006	rev 1.0
    	original version

    hm	29. feb 2008	rev 1.1
    	improved performance

    hm	6. jun. 2008	rev 1.2
    	changes type of input N from byte to int
    *)

END_FUNCTION

(* ---- BIT_TOGGLE_B.st ---- *)
FUNCTION BIT_TOGGLE_B
    (*http://www.oscat.de/images/OSCATBasic/oscat_basic333_en.pdf#page=214*)
    BIT_TOGGLE_B := SHL(BYTE#1, POS) XOR IN;

    (* revision history
    hm	18. oct. 2008	rev 1.0
    	original version

    *)

END_FUNCTION

(* ---- BIT_TOGGLE_DW.st ---- *)
FUNCTION BIT_TOGGLE_DW
    (*http://www.oscat.de/images/OSCATBasic/oscat_basic333_en.pdf#page=214*)
    BIT_TOGGLE_DW := SHL(DWORD#1, POS) XOR IN;

    (* revision history
    hm	18. oct. 2008	rev 1.0
    	original version

    *)

END_FUNCTION

(* ---- BIT_TOGGLE_W.st ---- *)
FUNCTION BIT_TOGGLE_W
    (*http://www.oscat.de/images/OSCATBasic/oscat_basic333_en.pdf#page=215*)
    BIT_TOGGLE_W := SHL(WORD#1, POS) XOR IN;

    (* revision history
    hm	18. oct. 2008	rev 1.0
    	original version

    *)

END_FUNCTION

(* ---- BUFFER_COMP.st ---- *)
FUNCTION BUFFER_COMP
    (*http://www.oscat.de/images/OSCATBasic/oscat_basic333_en.pdf#page=480*)
    (* search for first character match *)
    IF SIZE2 <= SIZE1 THEN
    	end := SIZE1 - SIZE2;
    	firstbyte := PT2[0];
    	FOR i := START TO end DO
    		IF PT1[i] = firstbyte THEN
    			(* first character matches, now compare rest of array *)
    			j := 1;
    			WHILE j < SIZE2 DO
    				IF PT2[j] <> PT1[j+i] THEN EXIT; END_IF
    				j := j + 1;
    			END_WHILE
    			(* when j > SIZE2 a match was found return the position i in buffer1 *)
    			IF j = SIZE2 THEN
    				BUFFER_COMP := i;
    				RETURN;
    			END_IF
    		END_IF
    	END_FOR
    END_IF
    BUFFER_COMP := -1;

    (*
    hm 14. nov. 2008	rev 1.0
    	original version

    hm	12. nov. 2009	rev 1.1
    	performance increase

    *)
END_FUNCTION

(* ---- BUFFER_SEARCH.st ---- *)
FUNCTION BUFFER_SEARCH
    (*http://www.oscat.de/images/OSCATBasic/oscat_basic333_en.pdf#page=481*)
    ps ACCESS ADR(STR);
    lx := LEN(STR);
    end := MIN(SIZE - lx, SIZE - 1);
    lx := lx - 1;
    FOR i := POS TO end DO
    	FOR k := 0 TO lx DO
    		IF IGN THEN chx := TO_UPPER(PT[i+k]); ELSE chx := PT[i+k]; END_IF
    		IF ps[k] <> chx THEN EXIT; END_IF
    	END_FOR
    	IF k > lx THEN
    		BUFFER_SEARCH := i;
    		RETURN;
    	END_IF
    END_FOR
    BUFFER_SEARCH := -1;

    (* revision History

    hm 5. mar. 2008	rev 1.0
    	original version

    hm	16. mar. 2008	rev 1.1
    	chaged type of input SIZE to uint

    hm	13. may. 2008	rev 1.2
    	changed type of pointer to array[1..32767]
    	changed SIZE of string to STRING_LENGTH

    hm	12. nov. 2009	rev 1.3
    	limit end to array SIZE

    hm	25. jan. 2011	rev 1.4
    	IGN = True will now ignore case
    	return -1 if nothing found
    *)
END_FUNCTION

(* ---- BUFFER_TO_STRING.st ---- *)
FUNCTION BUFFER_TO_STRING
    (*http://www.oscat.de/images/OSCATBasic/oscat_basic333_en.pdf#page=482*)
    ps ACCESS ADR(RETVAL);
    IF SIZE = 0 THEN RETURN; END_IF
    sta := MIN(START, SIZE -1);
    stp := MIN(STOP, SIZE -1);

    (* check for maximum string_length *)
    IF UINT_TO_INT(stp - sta + 1) >= STRING_LENGTH THEN
    	stp := sta + INT_TO_UINT(STRING_LENGTH) - 1;
    END_IF

    FOR i := sta TO stp DO
    	ps := PT[i];
    	ps ACCESS (ADR(ps) + 1);
    END_FOR

    (* terminate the string *)

    ps := 0;
    BUFFER_TO_STRING := TRUE;

    (* revision History
    hm 	5. mar. 2008	rev 1.0
    	original version

    hm	16. mar. 2008	rev 1.1
    	changed type of input SIZE to uint

    hm	13. may. 2008	rev 1.2
    	changed type of pointer to array[0..32767]
    	changed SIZE of string to STRING_LENGTH

    hm	12. jun. 2008	rev 1.3
    	check for pointer overrun
    	change input START and STOP to uint
    	added type conversions to avoid warnings under codesys 3.0

    hm	23. mar. 2009	rev 1.4
    	avoid writing to input STOP

    hm	12. nov. 2009 rev 1.5
    	limit START and STOP to SIZE -1

    *)
END_FUNCTION

(* ---- BYTE_OF_BIT.st ---- *)
FUNCTION BYTE_OF_BIT
    (*http://www.oscat.de/images/OSCATBasic/oscat_basic333_en.pdf#page=215*)
    BYTE_OF_BIT := SHL(SHL(SHL(SHL(SHL(SHL(SHL(BOOL_TO_BYTE(B7),1) OR BOOL_TO_BYTE(B6),1) OR BOOL_TO_BYTE(B5),1) OR BOOL_TO_BYTE(B4),1)
    	OR BOOL_TO_BYTE(B3),1) OR BOOL_TO_BYTE(B2),1) OR BOOL_TO_BYTE(B1),1) OR BOOL_TO_BYTE(B0);

    (* revision history

    hm	4. aug 2006		rev 1.0
    	original version

    hm	18. feb. 2008	rev 1.1
    	improved performance

    *)
END_FUNCTION

(* ---- BYTE_OF_DWORD.st ---- *)
FUNCTION BYTE_OF_DWORD
    (*http://www.oscat.de/images/OSCATBasic/oscat_basic333_en.pdf#page=216*)
    BYTE_OF_DWORD := DWORD_TO_BYTE(SHR(IN,SHL(N,3)));

    (* revision history
    hm	17. jan 2007	rev 1.0
    	original version

    hm	2. jan 2008		rev 1.1
    	improved performance

    hm	30. oct. 2008	rev 1.2
    	improved performance
    *)

END_FUNCTION

(* ---- BYTE_TO_GRAY.st ---- *)
FUNCTION BYTE_TO_GRAY
    (*http://www.oscat.de/images/OSCATBasic/oscat_basic333_en.pdf#page=217*)
    BYTE_TO_GRAY := IN XOR SHR(IN,1);

    (* revision history
    hm	9. nov. 2009	rev 1.0
    	original version

    *)
END_FUNCTION

(* ---- BYTE_TO_RANGE.st ---- *)
FUNCTION BYTE_TO_RANGE
    (*http://www.oscat.de/images/OSCATBasic/oscat_basic333_en.pdf#page=273*)
    BYTE_TO_RANGE := (HIGH - LOW) * BYTE_TO_USINT(X) / 255.0 + LOW;

    (* revision history
    hm	9. jan 2008		rev 1.0
    	original version

    *)

END_FUNCTION

(* ---- BYTE_TO_STRB.st ---- *)
FUNCTION BYTE_TO_STRB
    (*http://www.oscat.de/images/OSCATBasic/oscat_basic333_en.pdf#page=145*)
    (* pointer für die ausgabe ermitteln *)
    pt ACCESS ADR(RETVAL);
    (* die 8 ausgabecharacter ermitteln und schreiben *)
    FOR i := 1 TO 8 DO
    	pt := USINT_TO_BYTE(BOOL_TO_USINT(IN.7) + 48);
    	IN := SHL(IN,1);
    	pt ACCESS (ADR(pt) + 1);
    END_FOR

    (* der ausgabestring muss noch mit 0 abgeschlossen werden *)
    pt := 0;

    BYTE_TO_STRB := TRUE;

    (* code before rev 1.1
    FOR i := 1 TO 8 DO
    	IF IN.0 = 0 THEN temp := CONCAT('0', temp); ELSE temp := CONCAT('1', temp); END_IF
    	IN := SHR(IN, 1);
    END_FOR
    BYTE_TO_STRB := temp;
    *)

    (* revision history

    hm		9.6.2007	rev 1.0
    	original version

    hm	15. dec 2007	rev 1.1
    	inprooved code for higher performance

    hm	29. mar. 2008	rev 1.2
    	changed STRING to STRING(8)

    hm	20. jun. 2008	rev 1.3
    	performance improvement

    *)
END_FUNCTION

(* ---- BYTE_TO_STRH.st ---- *)
FUNCTION BYTE_TO_STRH
    (*http://www.oscat.de/images/OSCATBasic/oscat_basic333_en.pdf#page=146*)
    (* read pointer to output string *)
    PT ACCESS ADR(BYTE_TO_STRH);
    (* calculate high order hex value *)
    temp := SHR(IN,4);
    intTemp := BYTE_TO_USINT(temp);
    (* convert value to hex character *)
    IF intTemp <= 9 THEN temp := USINT_TO_BYTE(intTemp + 48); ELSE temp := USINT_TO_BYTE(intTemp + 55); END_IF
    (* write friat character to output string *)
    PT := temp;
    (* calculate low order hex value *)
    temp := IN AND 2#00001111;
    intTemp := BYTE_TO_USINT(temp);
    IF intTemp <= 9 THEN temp := USINT_TO_BYTE(intTemp + 48); ELSE temp := USINT_TO_BYTE(intTemp + 55); END_IF
    (* increment pointer and wirte low order character *)
    PT ACCESS (ADR(PT) + 1);
    PT := temp;
    (* set pointer at the end of the output string and close the string with 0 *)
    PT ACCESS (ADR(PT) + 1);
    PT:= 0;

    (* code before rev 1.2
    FOR i := 1 TO 2 DO
    	X := IN AND 2#1111;
    	IF X <= 9 THEN X := X + 48; ELSE X := X + 55; END_IF
    	Cx := CHR(X);
    	temp := CONCAT(Cx, temp);
    	IN := SHR(IN,4);
    END_FOR
    BYTE_TO_STRH := temp;
    *)

    (* revision history

    hm	9.6.2007		rev 1.0
    	original version

    hm	11.9.2007		rev 1.1
    	changed coding for compatibility with twincat, under twincat concat cannot have a function as argument.

    hm	15 dec 2007		REV 1.2
    	changed code for higher performance

    hm	29. mar. 2008	rev 1.3
    	changed STRING to STRING(2)
    *)
END_FUNCTION

(* ---- C_TO_F.st ---- *)
FUNCTION C_TO_F
    (*http://www.oscat.de/images/OSCATBasic/oscat_basic333_en.pdf#page=356*)
    C_TO_F := CELSIUS * 1.8 + 32.0;

    (* revision history

    hm	4. aug. 2006	rev 1.0
    	original version

    hm	11. mar. 2009	rev 1.1
    	real constants updated to new systax using dot

    *)
END_FUNCTION

(* ---- C_TO_K.st ---- *)
FUNCTION C_TO_K
    (*http://www.oscat.de/images/OSCATBasic/oscat_basic333_en.pdf#page=356*)
    C_TO_K := CELSIUS - cT0;

    (* revision history

    hm	4. aug 2006	rev 1.0
    	original version

    hm	19. aug 2009	rev 1.1
    	fixed calculation error

    *)

END_FUNCTION

(* ---- CABS.st ---- *)
FUNCTION CABS
    (*http://www.oscat.de/images/OSCATBasic/oscat_basic333_en.pdf#page=83*)
    CABS := HYPOT(X.re, X.im);

    (* revision history
    hm	21. feb 2008	rev 1.0
    	original version

    *)
END_FUNCTION

(* ---- CACOS.st ---- *)
FUNCTION CACOS
    (*http://www.oscat.de/images/OSCATBasic/oscat_basic333_en.pdf#page=83*)
    CACOSH(X,Y);
    RETVAL.re := Y.im;
    RETVAL.im := -Y.re;

    CACOS:=TRUE;

    (* revision history
    hm	21. feb 2008	rev 1.0
    	original version

    *)
END_FUNCTION

(* ---- CACOSH.st ---- *)
FUNCTION CACOSH
    (*http://www.oscat.de/images/OSCATBasic/oscat_basic333_en.pdf#page=84*)
    Y.re := (X.re - X.im)*(X.re + X.im) - 1.0;
    Y.im := 2.0 * X.re * X.im;
    CSQRT(Y, Y);
    Y.re := Y.re + X.re;
    Y.im := Y.im + X.im;
    CLOG(Y, RETVAL);
    CACOSH  := TRUE;

    (* revision history
    hm	21. feb 2008	rev 1.0
    	original version

    *)
END_FUNCTION

(* ---- CADD.st ---- *)
FUNCTION CADD
    (*http://www.oscat.de/images/OSCATBasic/oscat_basic333_en.pdf#page=84*)
    RETVAL.re := X.re + Y.re;
    RETVAL.im := X.im + Y.im;
    CADD:=TRUE;

    (* revision history
    hm	21. feb 2008	rev 1.0
    	original version

    *)
END_FUNCTION

(* ---- CAPITALIZE.st ---- *)
FUNCTION CAPITALIZE
    (*http://www.oscat.de/images/OSCATBasic/oscat_basic333_en.pdf#page=146*)
    PT ACCESS ADR(RETVAL);
    RETVAL := STR;
    L := LEN(STR);
    FOR pos := 1 TO L DO
    	IF first THEN PT := TO_UPPER(PT);	END_IF
    	(* remember in first if the next char needs to capitalized *)
    	first := PT= 32;
    	PT ACCESS (ADR(PT) + 1);
    END_FOR
    CAPITALIZE := TRUE;
    (* revision histroy
    hm		4. mar 2008	rev 1.0
    	original release

    hm	29. mar. 2008	rev 1.1
    	changed STRING to STRING(STRING_LENGTH)

    hm	20. jun. 2008	rev 1.2
    	improved performance

    *)

END_FUNCTION

(* ---- CARG.st ---- *)
FUNCTION CARG
    (*http://www.oscat.de/images/OSCATBasic/oscat_basic333_en.pdf#page=84*)
    CARG := ATAN2(X.im, X.re);

    (* revision history
    hm	21. feb. 2008	rev 1.0
    	original version

    hm	20. apr. 2008	rev 1.1
    	use ATAN2 instead of ATAN
    *)
END_FUNCTION

(* ---- CASIN.st ---- *)
FUNCTION CASIN
    (*http://www.oscat.de/images/OSCATBasic/oscat_basic333_en.pdf#page=85*)
    Y.re := -X.im;
    Y.im := X.re;
    CASINH(Y, Y);
    RETVAL.re := Y.im;
    RETVAL.im := -Y.re;
    CASIN := TRUE;

    (* revision history
    hm	21. feb 2008	rev 1.0
    	original version

    *)
END_FUNCTION

(* ---- CASINH.st ---- *)
FUNCTION CASINH
    (*http://www.oscat.de/images/OSCATBasic/oscat_basic333_en.pdf#page=85*)
    Y.re := (X.re - X.im)*(X.re + X.im) + 1.0;
    Y.im := 2.0 * X.re * X.im;
    CSQRT(Y,Y);
    Y.re := Y.re + X.re;
    Y.im := Y.im + X.im;
    CLOG(Y,RETVAL);
    CASINH  := TRUE;

    (* revision history
    hm	21. feb 2008	rev 1.0
    	original version

    *)
END_FUNCTION

(* ---- CATAN.st ---- *)
FUNCTION CATAN
    (*http://www.oscat.de/images/OSCATBasic/oscat_basic333_en.pdf#page=86*)
    r2 := X.re * X.re;
    den := 1.0 - r2 - X.im * X.im;
    RETVAL.re := 0.5 * ATAN(2.0 * X.re / den);
    num := X.im + 1.0;
    num := r2 + num * num;
    den := X.im - 1.0;
    den := r2 + den * den;
    RETVAL.im := 0.25 * (LN(num)-LN(den));
    CATAN:=TRUE;
    (* revision history
    hm	21. feb 2008	rev 1.0
    	original version

    *)
END_FUNCTION

(* ---- CATANH.st ---- *)
FUNCTION CATANH
    (*http://www.oscat.de/images/OSCATBasic/oscat_basic333_en.pdf#page=86*)
    i2 := X.im * X.im;
    num := 1.0 + X.re;
    num := i2 + num * num;
    den := 1.0 - X.re;
    den := i2 + den * den;
    RETVAL.re := 0.25 * (LN(num) - LN(den));
    den := 1 - X.re * X.re - i2;
    RETVAL.im := 0.5 * ATAN(2.0 * X.im / den);
    CATANH:=TRUE;
    (* revision history
    hm	21. feb 2008	rev 1.0
    	original version

    *)
END_FUNCTION

(* ---- CAUCHY.st ---- *)
FUNCTION CAUCHY
    (*http://www.oscat.de/images/OSCATBasic/oscat_basic333_en.pdf#page=42*)
    tmp := X - T;
    CAUCHY := cPI_INV * U / (U*U + tmp*tmp);

    (* revision hisdtory
    hm	26. oct. 2008	rev 1.0
    	original version

    *)
END_FUNCTION

(* ---- CAUCHYCD.st ---- *)
FUNCTION CAUCHYCD
    (*http://www.oscat.de/images/OSCATBasic/oscat_basic333_en.pdf#page=43*)
    CAUCHYCD := 0.5 + cPI_INV * ATAN((X - T) / U);

    (* revision hisdtory
    hm	26. oct. 2008	rev 1.0
    	original version

    *)
END_FUNCTION

(* ---- CCON.st ---- *)
FUNCTION CCON
    (*http://www.oscat.de/images/OSCATBasic/oscat_basic333_en.pdf#page=86*)
    RETVAL.re := X.re;
    RETVAL.im := -X.im;
    CCON:=TRUE;

    (* revision history
    hm	21. feb 2008	rev 1.0
    	original version

    *)
END_FUNCTION

(* ---- CCOS.st ---- *)
FUNCTION CCOS
    (*http://www.oscat.de/images/OSCATBasic/oscat_basic333_en.pdf#page=87*)
    CSET(-X.im, X.re, temp);
    CCOSH(temp,RETVAL);
    CCOS := TRUE;

    (* revision history
    hm	21. feb 2008	rev 1.0
    	original version

    *)
END_FUNCTION

(* ---- CCOSH.st ---- *)
FUNCTION CCOSH
    (*http://www.oscat.de/images/OSCATBasic/oscat_basic333_en.pdf#page=87*)
    RETVAL.re := COSH(X.re) * COS(X.im);
    RETVAL.im := SINH(X.re) * SIN(X.im);
    CCOSH := TRUE;

    (* revision history
    hm	21. feb 2008	rev 1.0
    	original version

    *)
END_FUNCTION

(* ---- CDIV.st ---- *)
FUNCTION CDIV
    (*http://www.oscat.de/images/OSCATBasic/oscat_basic333_en.pdf#page=87*)
    Temp := Y.re * Y.re + Y.im * Y.im;
    RETVAL.re := (X.re * Y.re + X.im * Y.im) / Temp;
    RETVAL.im := (X.im * Y.re - X.re * Y.im) / Temp;
    CDIV := TRUE;
    (* revision history
    hm	21. feb 2008	rev 1.0
    	original version

    *)
END_FUNCTION

(* ---- CEIL.st ---- *)
FUNCTION CEIL
    (*http://www.oscat.de/images/OSCATBasic/oscat_basic333_en.pdf#page=43*)
    CEIL := REAL_TO_INT(X);
    IF CEIL < X THEN
    	CEIL := CEIL + 1;
    END_IF

    (* revision history
    hm	7. feb. 2007	rev 1.0
    	original version

    hm	21. mar. 2008	rev 1.1
    	use REAL_TO_INT instead of trunc for compatibility reasons

    *)

END_FUNCTION

(* ---- CEIL2.st ---- *)
FUNCTION CEIL2
    (*http://www.oscat.de/images/OSCATBasic/oscat_basic333_en.pdf#page=44*)
    CEIL2 := REAL_TO_DINT(X);
    IF DINT_TO_REAL(CEIL2) < X THEN
    	CEIL2 := CEIL2 + 1;
    END_IF

    (* revision history
    hm	21. mar. 2008	rev 1.0
    	original version

    hm	4. apr. 2008	rev 1.1
    	added type conversion to avoid warnings under codesys 3.0

    hm	30. jun. 2008	rev 1.2
    	added type conversion to avoid warnings under codesys 3.0

    hm	10. mar. 2009	rev 1.3
    	use correct statement real_to_DINT

    *)

END_FUNCTION

(* ---- CEXP.st ---- *)
FUNCTION CEXP
    (*http://www.oscat.de/images/OSCATBasic/oscat_basic333_en.pdf#page=88*)
    Temp := EXP(X.re);
    RETVAL.re := Temp * COS(X.im);
    RETVAL.im := Temp * SIN(X.im);
    CEXP:=TRUE;

    (* revision history
    hm	21. feb 2008	rev 1.0
    	original version

    *)
END_FUNCTION

(* ---- CHARCODE.st ---- *)
FUNCTION CHARCODE
    (*http://www.oscat.de/images/OSCATBasic/oscat_basic333_en.pdf#page=147*)
    IF LEN(STR) = 1 THEN
    	CHARCODE := CODE(STR, 1);
    ELSIF STR <> '' THEN
    	(* construct search string *)
    	search := CONCAT('&', STR);
    	search := CONCAT(search, ';');
    	WHILE pos = 0 AND (i < 4) DO
    		i := i + 1;
    		pos := FIND(cCHARNAMES[i], search);
    	END_WHILE
    	found := MID(cCHARNAMES[i], 1, pos - 1);
    	CHARCODE := CODE(found, 1);
    END_IF

    (* revision history
    hm	13. may. 2008	rev 1.0
    	original version

    hm	19. oct. 2008	rev 1.1
    	changed setup constants

    hm	24. oct. 2008	rev 1.2
    	optimized code
    *)

END_FUNCTION

(* ---- CHARNAME.st ---- *)
FUNCTION CHARNAME
    (*http://www.oscat.de/images/OSCATBasic/oscat_basic333_en.pdf#page=147*)
    IF C <> 0 THEN
    	(* construct search string from code followed by $ sign, also clear CHARNAME string*)
    	CHR_TO_STRING(C, RETVAL);
    	RETVAL := CONCAT(RETVAL,'&');
    	RETVAL := CONCAT(';', RETVAL);
    	WHILE pos = 0 AND (i < 4) DO
    		i := i + 1;
    		pos := FIND(cCHARNAMES[i], RETVAL);
    	END_WHILE
    	IF pos > 0 THEN
    		RETVAL := MID(cCHARNAMES[i], 10, pos + 3);
    		(* search for end of name and truncate *)
    		pos := FIND(RETVAL, ';');
    		RETVAL := LEFT(RETVAL,pos - 1);
    	ELSE
    		 CHR_TO_STRING(C, RETVAL);
    	END_IF
        CHARNAME:=TRUE;
    ELSE
    	RETVAL := '';
        CHARNAME:=FALSE;
    END_IF

    (* revision history
    hm	13. may. 2008	rev 1.0
    	original version

    hm	16. jun. 2008	rev 1.1
    	changed nested call of concat for better compatibility

    hm	19. oct. 2008	rev 1.2
    	changes setup constants

    hm	24. oct. 2008	rev 1.3
    	new code for high performance

    hm	17. dec. 2008	rev 1.4
    	changed function chr to chr_to_string
    *)

END_FUNCTION

(* ---- CHECK_PARITY.st ---- *)
FUNCTION CHECK_PARITY
    (*http://www.oscat.de/images/OSCATBasic/oscat_basic333_en.pdf#page=217*)
    CHECK_PARITY := NOT P;
    WHILE IN > 0 DO
    	CHECK_PARITY := CHECK_PARITY XOR IN.0 XOR IN.1 XOR IN.2 XOR IN.3;
    	IN := SHR(IN,4);
    END_WHILE

    (* code before rev 1.2
    WHILE IN > 0 DO
    	IF IN.0 THEN cnt := cnt + 1; END_IF
    	IN := SHR(IN,1);
    END_WHILE
    CHECK_PARITY := even(cnt) XOR P;
    *)

    (* revision history

    rev 1.0 HM  1.oct.2006

    rev 1.1 hm	10.sep.2007
    	changed algorithm to improove performance

    rev 1.2	hm	8 dec 2007
    	changed algorithm to improove performance

    rev 1.3 hm	18. feb 2008
    	changed algorithm to improove performance
    *)
END_FUNCTION

(* ---- CHK_REAL.st ---- *)
FUNCTION CHK_REAL
    (*http://www.oscat.de/images/OSCATBasic/oscat_basic333_en.pdf#page=217*)
    pt ACCESS ADR(X);				(* move real to dword, real_to_dword does not work becasze it treats dword as a number on many systems *)
    tmp := ROL(pt,1);			(* rotate left foir easy checking, sign will be at lease significant digit *)
    IF DWORD_TO_UDINT(tmp) < 16#FF000000 THEN
    	CHK_REAL := 16#00;		(* normalized and denormalized numbers *)
    ELSIF tmp = 16#FF000000 THEN
    	CHK_REAL := 16#20;		(* X is +infinity see IEEE754 *)
    ELSIF tmp = 16#FF000001 THEN
    	CHK_REAL := 16#40;		(* X is -infinity see IEEE754 *)
    ELSE
    	CHK_REAL := 16#80;		(* X is NAN see IEEE754 *)
    END_IF

    (* revision history
    hm	 20. jan. 2011	rev 1.0
    	original version

    *)
END_FUNCTION

(* ---- CHR_TO_STRING.st ---- *)
FUNCTION CHR_TO_STRING
    (*http://www.oscat.de/images/OSCATBasic/oscat_basic333_en.pdf#page=148*)
    PT ACCESS ADR(RETVAL); //Assign the return value address to pointer
    PT := C; // set the pointers value to C
    PT ACCESS (ADR(PT) + 1); //increment the pointers value by one to get the next byte of the return string. STRING[1] is two bytes long
    PT := 0; //Set the pointer value to 0
    CHR_TO_STRING := TRUE;

    (* revision history
    hm	16 jan 2007		rev 1.0
    	original version

    hm	4. feb. 2008	rev 1.1
    	return string would not be terminated properly

    hm	29. mar. 2008	rev 1.2
    	changed STRING to STRING(1)

    hm	17. dec. 2008	rev 1.3
    	changed name of function from chr to CHR_TO_STRING
    *)
END_FUNCTION

(* ---- CINV.st ---- *)
FUNCTION CINV
    (*http://www.oscat.de/images/OSCATBasic/oscat_basic333_en.pdf#page=88*)
    temp := X.re * X.re + X.im * X.im;
    RETVAL.re := X.re / temp;
    RETVAL.im := -X.im / temp;
    CINV:=TRUE;
    (* revision history
    hm	21. feb 2008	rev 1.0
    	original version

    *)
END_FUNCTION

(* ---- CIRCLE_A.st ---- *)
FUNCTION CIRCLE_A
    (*http://www.oscat.de/images/OSCATBasic/oscat_basic333_en.pdf#page=104*)
    CIRCLE_A := RX * RX * 8.726646E-3 * AX;

    (* revision histroy
    hm	16. oct 2007	rev 1.0
    	original version

    hm	4. dec 2007		rev 1.1
    	changed code for better performance

    hm	22. feb 2008	rev 1.2
    	improved performance
    *)
END_FUNCTION

(* ---- CIRCLE_C.st ---- *)
FUNCTION CIRCLE_C
    (*http://www.oscat.de/images/OSCATBasic/oscat_basic333_en.pdf#page=104*)
    CIRCLE_C := 1.7453293E-2 * RX * AX;

    (* revision histroy
    hm	16. oct 2007	rev 1.0
    	original version

    hm	22. feb 2008	rev 1.1
    	improved performance
    *)
END_FUNCTION

(* ---- CIRCLE_SEG.st ---- *)
FUNCTION CIRCLE_SEG
    (*http://www.oscat.de/images/OSCATBasic/oscat_basic333_en.pdf#page=105*)
    IF RX > 0.0 THEN
    	CIRCLE_SEG := 2.0 * ACOS(1.0 - LIMIT(0.0, HX / RX, 2.0));
    	CIRCLE_SEG := (CIRCLE_SEG - SIN(CIRCLE_SEG)) *RX * RX / 2.0;
    END_IF

    (* revision histroy
    hm	10. mar 2010	rev 1.0
    	original version

    *)
END_FUNCTION

(* ---- CLEAN.st ---- *)
FUNCTION CLEAN
    (*http://www.oscat.de/images/OSCATBasic/oscat_basic333_en.pdf#page=149*)
    (* copy input string *)
    RETVAL := IN;
    stop := LEN(IN);
    WHILE pos <= stop DO
    	IF FIND(CX, MID(RETVAL, 1, pos)) > 0 THEN
    		(* charcter found skip to next one *)
    		pos := pos + 1;
    	ELSE
    		(* wrong chracter needs to be deleted *)
    		RETVAL := DELETE(RETVAL, 1, pos);
    		stop := stop - 1;	(* the string is one character shorter now *)
    	END_IF
    END_WHILE
    CLEAN := TRUE;

    (* revision history

    hm		18. jun. 2008	rev 1.0
    	original version

    *)
END_FUNCTION

(* ---- CLOG.st ---- *)
FUNCTION CLOG
    (*http://www.oscat.de/images/OSCATBasic/oscat_basic333_en.pdf#page=88*)
    RETVAL.re := LN(HYPOT(X.re, X.im));
    RETVAL.im := ATAN2(X.im, X.re);
    CLOG := TRUE;

    (* revision history
    hm	21. feb 2008	rev 1.0
    	original version

    hm	20. apr. 2008	rev 1.1
    	use ATAN2 instead of ATAN
    *)
END_FUNCTION

(* ---- CMP.st ---- *)
FUNCTION CMP
    (*http://www.oscat.de/images/OSCATBasic/oscat_basic333_en.pdf#page=44*)
    tmp := ABS(X);
    IF tmp > 0.0 THEN
    	tmp := EXP10(INT_TO_REAL(FLOOR(LOG(tmp))-N+1));
    ELSE
    	tmp := EXP10(tmp);
    END_IF
    CMP := ABS(X - Y) < tmp;

    (* revision history
    hm	12. mar. 2008	rev 1.0
    	original version

    hm	10. mar. 2009	rev 1.1
    	added type conversion for compatibility reasons
    *)

END_FUNCTION

(* ---- CMUL.st ---- *)
FUNCTION CMUL
    (*http://www.oscat.de/images/OSCATBasic/oscat_basic333_en.pdf#page=89*)
    RETVAL.re := X.re * Y.re - X.im * Y.im;
    RETVAL.im := X.re * Y.im + X.im * Y.re;
    CMUL:=TRUE;
    (* revision history
    hm	21. feb 2008	rev 1.0
    	original version

    *)
END_FUNCTION

(* ---- CODE.st ---- *)
FUNCTION CODE
    (*http://www.oscat.de/images/OSCATBasic/oscat_basic333_en.pdf#page=149*)
    IF POS < 1 OR POS > LEN(STR) THEN
    	CODE := 0;
    	RETURN;
    ELSE
    	PT ACCESS (ADR(STR) + POS - 1);
    	CODE := PT;
    END_IF

    (* revision history
    hm	9. mar. 2008	rev 1.0
    	original version

    hm	29. mar. 2008	rev 1.1
    	changed STRING to STRING(STRING_LENGTH)
    *)
END_FUNCTION

(* ---- CONE_V.st ---- *)
FUNCTION CONE_V
    (*http://www.oscat.de/images/OSCATBasic/oscat_basic333_en.pdf#page=105*)
    CONE_V := 1.047197551 * RX * RX * HX;

    (* revision histroy
    hm	17. oct 2007	rev 1.0
    	original version

    hm	4. dec 2007		rev 1.1
    	changed code for better performance

    hm	22. feb 2008	rev 1.2
    	changed code for better performance
    *)
END_FUNCTION

(* ---- COSH.st ---- *)
FUNCTION COSH
    (*http://www.oscat.de/images/OSCATBasic/oscat_basic333_en.pdf#page=45*)
    t := EXP(X);
    COSH := (1.0 / t + t) * 0.5;

    (* revision histroy
    hm	12.1.2007	rev 1.0
    	original version

    hm	1.12.2007	rev 1.1
    	changed code to improve performance

    hm	5. jan 2008	rev 1.2
    	further performance improvement

    hm	10. mar. 2009	rev 1.3
    	real constants updated to new systax using dot
    *)
END_FUNCTION

(* ---- COTH.st ---- *)
FUNCTION COTH
    (*http://www.oscat.de/images/OSCATBasic/oscat_basic333_en.pdf#page=45*)
    IF X > 20.0 THEN
    	COTH :=1.0;
    ELSIF X < -20.0 THEN
    	COTH := -1.0;
    ELSE
    	COTH := 1.0 + 2.0 / (EXP(X * 2.0) - 1.0);
    END_IF

    (* revision histroy
    hm		12.1.2007	rev 1.0
    	original version

    hm	1.12.2007		rev 1.1
    	changed code to improve performance

    hm	8. jan 2008	rev 1.2
    	further improvement in performance

    hm	10. mar 2008	rev 1.3
    	extended range of valid inputs to +/- INV
    	changed formula for better accuracy

    hm	10. mar. 2009	rev 1.4
    	real constants updated to new systax using dot
    *)
END_FUNCTION

(* ---- COUNT_CHAR.st ---- *)
FUNCTION COUNT_CHAR
    (*http://www.oscat.de/images/OSCATBasic/oscat_basic333_en.pdf#page=150*)
    pt ACCESS ADR(STR);
    l := LEN(STR);
    COUNT_CHAR := 0;
    FOR pos := 1 TO l DO
    	IF pt = CHR THEN COUNT_CHAR := COUNT_CHAR + 1; END_IF
        pt ACCESS (ADR(pt) + 1);
    END_FOR

    (* revision history
    hm	29. feb 2008	rev 1.0
    	original version

    hm	29. mar. 2008	rev 1.1
    	changed STRING to STRING(STRING_LENGTH)
    *)
END_FUNCTION

(* ---- COUNT_SUBSTRING.st ---- *)
FUNCTION COUNT_SUBSTRING
    (*http://www.oscat.de/images/OSCATBasic/oscat_basic333_en.pdf#page=150*)
    COUNT_SUBSTRING := 0;
    size := LEN(SEARCH);
    REPEAT
       pos := FIND(STR,SEARCH);
       IF pos > 0 THEN
          STR := REPLACE(STR, '', size,pos);
          COUNT_SUBSTRING := COUNT_SUBSTRING + 1;
       END_IF
    UNTIL pos = 0
    END_REPEAT

    (* revision history
    ks	20. jan. 2011	rev 1.0
    	original version

    *)

END_FUNCTION

(* ---- CPOL.st ---- *)
FUNCTION CPOL
    (*http://www.oscat.de/images/OSCATBasic/oscat_basic333_en.pdf#page=89*)
    RETVAL.re := L * COS(A);
    RETVAL.im := L * SIN(A);
    CPOL:=TRUE;

    (* revision history
    hm	21. feb 2008	rev 1.0
    	original version

    *)
END_FUNCTION

(* ---- CPOW.st ---- *)
FUNCTION CPOW
    (*http://www.oscat.de/images/OSCATBasic/oscat_basic333_en.pdf#page=89*)
    CLOG(X,temp);
    CMUL(Y,temp, temp2);
    CEXP(temp2, RETVAL);
    CPOW := TRUE;

    (* revision history
    hm	21. feb 2008	rev 1.0
    	original version

    *)
END_FUNCTION

(* ---- CRC_GEN.st ---- *)
FUNCTION CRC_GEN
    (*http://www.oscat.de/images/OSCATBasic/oscat_basic333_en.pdf#page=219*)
    (* align polygon *)
    shift := 32 - PL;
    PN := SHL(PN, shift);

    (* load first 4 bytes into register minimum message SIZE is 4 bytes
    	for smaller messages fill with 0#s at the beginning*)
    FOR pos := 0 TO 3 DO
    	IF REV_IN THEN CRC_GEN := SHL(CRC_GEN, 8) OR REVERSE(PT[pos]); ELSE CRC_GEN := SHL(CRC_GEN, 8) OR PT[pos]; END_IF
    END_FOR
    pos := 4;

    (* xor with INIT value *)
    CRC_GEN := CRC_GEN XOR SHL(INIT, shift);

    (* calculate CRC for each byte *)
    WHILE pos < SIZE DO
    	IF REV_IN THEN dx := REVERSE(PT[pos]); ELSE dx := PT[pos]; END_IF
    	pos := pos + 1;
    	(* crc calculation for one byte *)
    	FOR bits := 0 TO 7 DO
    		IF CRC_GEN.31 THEN
    			CRC_GEN := (SHL(CRC_GEN, 1) OR BOOL_TO_DWORD(dx.7)) XOR PN;
    		ELSE
    			CRC_GEN := SHL(CRC_GEN, 1) OR BOOL_TO_DWORD(dx.7);
    		END_IF
    		dx := SHL(dx, 1);
    	END_FOR
    END_WHILE

    (* all bytes are processed, need to finish the registers 32 bits *)
    FOR bits := 0 TO 31 DO
    	IF CRC_GEN.31 THEN
    		CRC_GEN := (SHL(CRC_GEN, 1) ) XOR PN;
    	ELSE
    		CRC_GEN := SHL(CRC_GEN, 1);
    	END_IF
    END_FOR

    (* final XOR *)
    CRC_GEN := SHR(CRC_GEN, shift) XOR XOR_OUT;

    (* reverse the crc_out put if necessary *)
    IF REV_OUT THEN CRC_GEN := REFLECT(CRC_GEN, PL); END_IF

    (* suggested optimization by deninis klopke
    die betreffs genannte Funktion kann folgendermaßen optimiert werden:
    In Zeilen 33 und 35 des Implementierungsteils kann jeweils der Teil „OR BOOL_TO_DWORD(dx.7)“ entfallen, da nach 8maligem Linksshift von „dx“ in Zeile 26 der Wert von dx = BYTE#0 ist. Eine weitere Veroderung mit diesem Wert hat keine Auswirkungen auf das Ergebnis mehr.
    *)

    (* typical crc polynoms

    CRC-4-ITU 			x4 + x + 1 					(ITU G.704, p. 12) 	0x3 or 0xC (0x9)
    CRC-5-ITU 			x5 + x4 + x2 + 1 			(ITU G.704, p. 9) 	0x15 or 0x15 (0x0B) Bluetooth
    CRC-5-USB 			x5 + x2 + 1 				(use: USB token packets) 	0x05 or 0x14 (0x9)
    CRC-6-ITU 			x6 + x + 1 					(ITU G.704, p. 3) 	0x03 or 0x30 (0x21)
    CRC-7 				x7 + x3 + 1 				(use: telecom systems, MMC) 	0x09 or 0x48 (0x11)
    CRC-8-ATM 			x8 + x2 + x + 1 				(use: ATM HEC) 	0x07 or 0xE0 (0xC1)
    CRC-8-CCITT 		x8 + x7 + x3 + x2 + 1 		(use: 1-Wire bus) 	0x8D or 0xB1 (0x63)
    CRC-8-Dallas/Maxim 	x8 + x5 + x4 + 1 			(use: 1-Wire bus) 	0x31 or 0x8C (0x19)
    CRC-8 				x8 + x7 + x6 + x4 + x2 + 1 	0xD5 or 0xAB (0x57)
    CRC-8-SAE J1850 	x8 + x4 + x3 + x2 + 1 		0x1D or 0xB8
    CRC-10 				x10 + x9 + x5 + x4 + x + 1 	0x233 or 0x331 (0x263)
    CRC-12 				x12 + x11 + x3 + x2 + x + 1 (use: telecom systems) 	0x80F or 0xF01 (0xE03)
    CRC-15-CAN 			x15 + x14 + x10 + x8 + x7 + x4 + x3 + 1 	0x4599 or 0x4CD1 (0x19A3)
    CRC-16-Fletcher 	Not a CRC; see Fletcher's checksum 	Used in Adler-32 A & B CRCs
    CRC-16-CCITT 	x16 + x12 + x5 + 1 (XMODEM,X.25, V.41, Bluetooth, PPP, IrDA; known as "CRC-CCITT") 	0x1021 or 0x8408 (0x0811)
    CRC-16-IBM 	x16 + x15 + x2 + 1 (USB, many others; also known as "CRC-16") 	0x8005 or 0xA001 (0x4003)
    CRC-24-Radix-64 	x24 + x23 + x18 + x17 + x14 + x11 + x10 + x7 + x6 + x5 + x4 + x3 + x + 1 	0x864CFB or 0xDF3261 (0xBE64C3)
    CRC-32-Adler 	Not a CRC; see Adler-32 	See Adler-32
    CRC-32-MPEG2 	x32 + x26 + x23 + x22 + x16 + x12 + x11 + x10 + x8 + x7 + x5 + x4 + x2 + x + 1 	0x04C11DB7 or 0xEDB88320 (0xDB710641) Also used in IEEE 802.3
    CRC-32-IEEE 802.3 	x32 + x26 + x23 + x22 + x16 + x12 + x11 + x10 + x8 + x7 + x5 + x4 + x2 + x + 1 (V.42) 	0x04C11DB7 or 0xEDB88320 (0xDB710641)
    CRC-32C (Castagnoli) 	x32 + x28 + x27 + x26 + x25 + x23 + x22 + x20 + x19 + x18 + x14 + x13 + x11 + x10 + x9 + x8 + x6 + 1 	0x1EDC6F41 or 0x82F63B78 (0x05EC76F1)
    CRC-64-ISO 	x64 + x4 + x3 + x + 1 (use: ISO 3309) 	0x000000000000001B or 0xD800000000000000 (0xB000000000000001)
    CRC-64-ECMA-182 	x64 + x62 + x57 + x55 + x54 + x53 + x52 + x47 + x46 + x45 + x40 + x39 + x38 + x37 + x35 + x33 + x32 + x31 + x29 + x27 + x24 + x23 + x22 + x21 + x19 + x17 + x13 + x12 + x10 + x9 + x7 + x4 + x + 1
    (as described in ECMA-182 p.63) 	0x42F0E1EBA9EA3693 or 0xC96C5795D7870F42 (0x92D8AF2BAF0E1E85)
    *)

    (* revision history

    hm	9.6.2007		rev 1.0
    	original version

    hm	11.9.2007		rev 1.1
    	deleted unused variable i

    hm	9. oct 2007 	rev 1.2
    	added INIT code for crc and XOR_OUT
    	added refelct in and reflect_out (REV_IN und REV_OUT)

    hm	2. jan 2008	rev 1.3
    	small changes for performance improvements

    hm	16. mar. 2008	rev 1.4
    	changed type of input SIZE to uint

    hm	10. mar. 2009	rev 1.5
    	removed nested comments

    hm	16. jan. 2011	rev 2.0
    	new version

    dk 3. feb 2021		rev 2.1
    	improved code by dennis koepke

    *)
END_FUNCTION

(* ---- CSET.st ---- *)
FUNCTION CSET
    (*http://www.oscat.de/images/OSCATBasic/oscat_basic333_en.pdf#page=90*)
    RETVAL.re := RE;
    RETVAL.im := IM;
    CSET:=TRUE;
    (* revision history
    hm	21. feb 2008	rev 1.0
    	original version

    *)
END_FUNCTION

(* ---- CSIN.st ---- *)
FUNCTION CSIN
    (*http://www.oscat.de/images/OSCATBasic/oscat_basic333_en.pdf#page=90*)
    RETVAL.re := COSH(X.im) * SIN(X.re);
    RETVAL.im := SINH(X.im) * COS(X.re);
    CSIN:=TRUE;

    (* revision history
    hm	21. feb 2008	rev 1.0
    	original version

    *)
END_FUNCTION

(* ---- CSINH.st ---- *)
FUNCTION CSINH
    (*http://www.oscat.de/images/OSCATBasic/oscat_basic333_en.pdf#page=90*)
    RETVAL.re := SINH(X.re) * COS(X.im);
    RETVAL.im := COSH(X.re) * SIN(X.im);
    CSINH:=TRUE;

    (* revision history
    hm	21. feb 2008	rev 1.0
    	original version

    *)
END_FUNCTION

(* ---- CSQRT.st ---- *)
FUNCTION CSQRT
    (*http://www.oscat.de/images/OSCATBasic/oscat_basic333_en.pdf#page=91*)
    temp := HYPOT(X.re, X.im);
    RETVAL.re :=  SQRT(0.5 * (temp + X.re));
    RETVAL.im :=  SGN(X.im) * SQRT(0.5 * (temp - X.re));
    CSQRT:=TRUE;

    (* revision history
    hm	21. feb 2008	rev 1.0
    	original version

    *)
END_FUNCTION

(* ---- CSUB.st ---- *)
FUNCTION CSUB
    (*http://www.oscat.de/images/OSCATBasic/oscat_basic333_en.pdf#page=91*)
    RETVAL.re := X.re - Y.re;
    RETVAL.im := X.im - Y.im;
    CSUB:=TRUE;
    (* revision history
    hm	21. feb 2008	rev 1.0
    	original version

    *)
END_FUNCTION

(* ---- CTAN.st ---- *)
FUNCTION CTAN
    (*http://www.oscat.de/images/OSCATBasic/oscat_basic333_en.pdf#page=91*)
    xi2 := 2.0 * X.im;
    xr2 := 2.0 * X.re;
    temp := 1.0 / (COS(xr2) + COSH( xi2));
    RETVAL.re := temp * SIN(xr2);
    RETVAL.im := temp * SINH(xi2);
    CTAN:=TRUE;

    (* revision history
    hm	21. feb 2008	rev 1.0
    	original version

    hm	10. mar 2009	rev 1.1
    	faster code
    *)
END_FUNCTION

(* ---- CTANH.st ---- *)
FUNCTION CTANH
    (*http://www.oscat.de/images/OSCATBasic/oscat_basic333_en.pdf#page=92*)
    xi2 := 2.0 * X.im;
    xr2 := 2.0 * X.re;
    temp := 1.0 / (COSH(xr2) + COS(xi2));
    RETVAL.re := temp * SINH(xr2);
    RETVAL.im := temp * SIN(xi2);
    CTANH:=TRUE;

    (* revision history
    hm	21. feb 2008	rev 1.0
    	original version

    hm	10. mar. 2009	rev 1.1
    	new faster code

    *)
END_FUNCTION

(* ---- CTRL_IN.st ---- *)
FUNCTION CTRL_IN
    (*http://www.oscat.de/images/OSCATBasic/oscat_basic333_en.pdf#page=380*)
    (* calculate the process error DIFF *)
    CTRL_IN := DEAD_ZONE(SET_POINT - ACTUAL, NOISE);

    (* revision history
    hm 	2. jun. 2008 	rev 1.0
    	original version

    *)
END_FUNCTION

(* ---- D_TRUNC.st ---- *)
FUNCTION D_TRUNC
    (*http://www.oscat.de/images/OSCATBasic/oscat_basic333_en.pdf#page=46*)
    D_TRUNC := REAL_TO_DINT(X);
    IF X > 0.0 THEN
    	IF DINT_TO_REAL(D_TRUNC) > X THEN D_TRUNC := D_TRUNC - 1; END_IF
    ELSE
    	IF DINT_TO_REAL(D_TRUNC) < X THEN D_TRUNC := D_TRUNC + 1; END_IF
    END_IF

    (* for systems that support a dint truncation this routine can be replaced by trunc() *)

    (* revision history
    hm	21. mar. 2008	rev 1.0
    	original version

    hm	31. oct. 2008	rev 1.1
    	optimized performance

    hm	10. mar. 2009	rev 1.2
    	real constants updated to new systax using dot
    *)
END_FUNCTION

(* ---- DATE_ADD.st ---- *)
FUNCTION DATE_ADD
    (*http://www.oscat.de/images/OSCATBasic/oscat_basic333_en.pdf#page=115*)
    DATE_ADD := UDINT_TO_DATE(DATE_TO_UDINT(IDATE) + INT_TO_UDINT(D + W * 7) * UDINT#86400);
    yr := Y + YEAR_OF_DATE(DATE_ADD);
    mo := M + MONTH_OF_DATE(DATE_ADD);
    dm := DAY_OF_MONTH(DATE_ADD);
    WHILE mo > 12 DO
    	mo := mo - 12;
    	yr := yr + 1;
    END_WHILE
    WHILE mo < 1 DO
    	mo := mo + 12;
    	yr := yr - 1;
    END_WHILE
    DATE_ADD := SET_DATE(yr, mo, dm);

    (* revision history

    hm 27.12.2006	rev 1.0
    	nrw module

    hm 12.4.2007		rev 1.1
    	corrected an error while date would be incorrect when year  = 0

    hm	1.11.2007		rev 1.2
    	added int_to_dword stetements to avoid possible overrun with möller ecp4

    hm	22. mar. 2008	rev 1.3
    	fixed some bugs when month was negative

    hm	7. oct. 2008	rev 1.4
    	changed function year to year_of_date
    	changed function month to month_of_date

    hm	29. mar. 2009	rev 1.5
    	improved performance

    hm	27. jan. 2011	rev 1.6
    	faster code

    hm	2. feb. 2011		rev 1.7
    	fixed an error, weeks not calculated

    hm	22. mar. 2011	rev 1.8
    	fixed an error in formula
    *)
END_FUNCTION

(* ---- DAY_OF_DATE.st ---- *)
FUNCTION DAY_OF_DATE
    (*http://www.oscat.de/images/OSCATBasic/oscat_basic333_en.pdf#page=116*)
    DAY_OF_DATE := UDINT_TO_DINT(DATE_TO_UDINT(IDATE) / 86400);

    (* revision history
    hm		16.9.2007		rev 1.0
    	original version

    hm		1. okt 2007		rev 1.1
    	added step7 compatibility

    hm		22. mar. 2008	rev 1.2
    	changed output from int to Dint because the total date range is 49710 days

    hm		7. apr. 2008	rev 1.3
    	deleted unused step7 code

    *)
END_FUNCTION

(* ---- DAY_OF_MONTH.st ---- *)
FUNCTION DAY_OF_MONTH
    (*http://www.oscat.de/images/OSCATBasic/oscat_basic333_en.pdf#page=116*)
    (* calculate the day in the year *)
    DAY_OF_MONTH := DAY_OF_YEAR(IDATE);
    (* leap will be set to one for a leap year *)
    leap := BOOL_TO_INT(LEAP_OF_DATE(IDATE));
    (* if leap year deduct one from the days of the year *)
    DAY_OF_MONTH := DAY_OF_MONTH - leap;
    (* search if we are in month december to march ? *)
    IF DAY_OF_MONTH > cMTH_OFS[9] THEN
    	IF DAY_OF_MONTH > cMTH_OFS[11] THEN
    		IF DAY_OF_MONTH > cMTH_OFS[12] THEN
    			DAY_OF_MONTH := DAY_OF_MONTH - cMTH_OFS[12];
    		ELSE
    			DAY_OF_MONTH := DAY_OF_MONTH - cMTH_OFS[11];
    		END_IF
    	ELSE
    		IF DAY_OF_MONTH > cMTH_OFS[10] THEN
    			DAY_OF_MONTH := DAY_OF_MONTH - cMTH_OFS[10];
    		ELSE
    			DAY_OF_MONTH := DAY_OF_MONTH - cMTH_OFS[9];
    		END_IF
    	END_IF
    ELSIF DAY_OF_MONTH > cMTH_OFS[5] THEN
    	IF DAY_OF_MONTH > cMTH_OFS[7] THEN
    		IF DAY_OF_MONTH > cMTH_OFS[8] THEN
    			DAY_OF_MONTH := DAY_OF_MONTH - cMTH_OFS[8];
    		ELSE
    			DAY_OF_MONTH := DAY_OF_MONTH - cMTH_OFS[7];
    		END_IF
    	ELSE
    		IF DAY_OF_MONTH > cMTH_OFS[6] THEN
    			DAY_OF_MONTH := DAY_OF_MONTH - cMTH_OFS[6];
    		ELSE
    			DAY_OF_MONTH := DAY_OF_MONTH - cMTH_OFS[5];
    		END_IF
    	END_IF
    ELSIF DAY_OF_MONTH > cMTH_OFS[3] THEN
    	IF DAY_OF_MONTH > cMTH_OFS[4] THEN
    		DAY_OF_MONTH := DAY_OF_MONTH - cMTH_OFS[4];
    	ELSE
    		DAY_OF_MONTH := DAY_OF_MONTH - cMTH_OFS[3];
    	END_IF
    ELSE
    	(* since now we must be in february or january we need to add leap again *)
    	DAY_OF_MONTH := DAY_OF_MONTH + leap;
    	IF DAY_OF_MONTH > cMTH_OFS[2] THEN DAY_OF_MONTH := DAY_OF_MONTH - cMTH_OFS[2]; END_IF
    	(* since nothing was true before, DAY_OF_MONTH must already be good *)
    END_IF

    (*
    Revision history

    hm 22.1.2007		rev 1.1
    	deleted unused variable day_in_year and day_in_year_begin

    hm	1. okt 2007	rev 1.2
    	changed code to use day_of_year and leap_of_date
    	added compatibility to STEP7

    hm	8. oct 2007	rev 1.3
    	deleted unused variable yr

    hm	8. jan 2008	rev 1.4
    	improved performance

    hm	25. oct. 2008	rev 2.0
    	new code using setup constants

    hm	10. mar. 2009	rev 2.1
    	removed nested comments

    *)

END_FUNCTION

(* ---- DAY_OF_WEEK.st ---- *)
FUNCTION DAY_OF_WEEK
    (*http://www.oscat.de/images/OSCATBasic/oscat_basic333_en.pdf#page=117*)
    DAY_OF_WEEK := UDINT_TO_INT((DATE_TO_UDINT(IDATE) / 86400 + 3) MOD 7) + 1;

    (* revision history
    hm 	21.8.06 		rev 1.1
    	corrected a miscalculation

    hm	23.12.2007		rev 1.2
    	correction for step7

    hm	7. apr. 2008	rev 1.3
    	deleted unused step7 code

    hm	7. oct. 2008	rev 1.4
    	changed name of function from weekday to DAY_OF_WEEK

    *)

END_FUNCTION

(* ---- DAY_OF_YEAR.st ---- *)
FUNCTION DAY_OF_YEAR
    (*http://www.oscat.de/images/OSCATBasic/oscat_basic333_en.pdf#page=117*)
    DAY_OF_YEAR := UDINT_TO_INT((DATE_TO_UDINT(IDATE) / UDINT#86400) MOD UDINT#1461);
    IF DAY_OF_YEAR > 729 THEN
    	IF DAY_OF_YEAR > 1095 THEN DAY_OF_YEAR := DAY_OF_YEAR - 1095; ELSE DAY_OF_YEAR := DAY_OF_YEAR - 729; END_IF
    ELSIF DAY_OF_YEAR > 364 THEN
    	DAY_OF_YEAR := DAY_OF_YEAR - 364;
    ELSE
    	DAY_OF_YEAR := DAY_OF_YEAR + 1;
    END_IF

    (*
    DAY_OF_YEAR := DWORD_TO_INT((DATE_TO_DWORD(IDATE) - DATE_TO_DWORD(YEAR_BEGIN(YEAR_OF_DATE(IDATE)))) / 86400) + 1;
    *)

    (* revivision history
    hm	4. aug. 2007		rev 1.0
    	original version

    hm	1. oct. 2007		rev 1.1
    	added compatibility to STEP7

    hm	4. jan. 2008		rev 1.2
    	changed code for better performance

    hm	7. oct. 2008		rev 1.3
    	changed name of function year to year_of_date

    hm	28. jan. 2011	rev 1.4
    	improved code
    *)
END_FUNCTION

(* ---- DAY_TO_TIME.st ---- *)
FUNCTION DAY_TO_TIME
    (*http://www.oscat.de/images/OSCATBasic/oscat_basic333_en.pdf#page=118*)
    DAY_TO_TIME := DWORD_TO_TIME(REAL_TO_DWORD(IN * 86400000.0));

    (* revision history
    hm	4. aug. 2006	rev 1.0
    	original release

    hm	24. feb. 2009	rev 1.1
    	renamed input to IN
    *)
END_FUNCTION

(* ---- DAYS_DELTA.st ---- *)
FUNCTION DAYS_DELTA
    (*http://www.oscat.de/images/OSCATBasic/oscat_basic333_en.pdf#page=118*)
    IF DATE_1 > DATE_2 THEN
    	DAYS_DELTA := - UDINT_TO_DINT((DATE_TO_UDINT(DATE_1) - DATE_TO_UDINT(DATE_2)) / 86400);
    ELSE
    	DAYS_DELTA := UDINT_TO_DINT((DATE_TO_UDINT(DATE_2) - DATE_TO_UDINT(DATE_1)) / 86400);
    END_IF

    (* revision history
    hm	27. dec 2006	rev 1.0
    	original version

    hm	16.9.2007		rev 1.1
    	coorected an error in formula and changed algorithm to show positive and negative delta

    hm	22. mar. 2008	rev 1.2
    	changed output from int to dint because the total date range is 49710 days

    hm	25. jan. 2011	rev 1.3
    	improved performance
    *)
END_FUNCTION

(* ---- DAYS_IN_MONTH.st ---- *)
FUNCTION DAYS_IN_MONTH
    (*http://www.oscat.de/images/OSCATBasic/oscat_basic333_en.pdf#page=119*)
    DAYS_IN_MONTH := DAY_OF_YEAR(IDATE);
    IF LEAP_OF_DATE(IDATE) THEN
    	CASE DAYS_IN_MONTH OF
    		32..60	:	DAYS_IN_MONTH := 29;
    		92..121 :	DAYS_IN_MONTH := 30;
    		153..182:	DAYS_IN_MONTH := 30;
    		245..274:	DAYS_IN_MONTH := 30;
    		306..335:	DAYS_IN_MONTH := 30;
    	ELSE
    		DAYS_IN_MONTH := 31;
    	END_CASE
    ELSE
    	CASE DAYS_IN_MONTH OF
    		32..59	:	DAYS_IN_MONTH := 28;
    		91..120 :	DAYS_IN_MONTH := 30;
    		152..181:	DAYS_IN_MONTH := 30;
    		244..273:	DAYS_IN_MONTH := 30;
    		305..334:	DAYS_IN_MONTH := 30;
    	ELSE
    		DAYS_IN_MONTH := 31;
    	END_CASE
    END_IF

    (* revision history
    hm	27. mar. 2009		rev 1.0
    	original version

    *)
END_FUNCTION

(* ---- DAYS_IN_YEAR.st ---- *)
FUNCTION DAYS_IN_YEAR
    (*http://www.oscat.de/images/OSCATBasic/oscat_basic333_en.pdf#page=119*)
    IF LEAP_OF_DATE(IDATE) THEN
    	DAYS_IN_YEAR := 366;
    ELSE
    	DAYS_IN_YEAR := 365;
    END_IF

    (* revision history
    hm	27. mar. 2009		rev 1.0
    	original version

    *)
END_FUNCTION

(* ---- DEAD_BAND.st ---- *)
FUNCTION DEAD_BAND
    (*http://www.oscat.de/images/OSCATBasic/oscat_basic333_en.pdf#page=387*)
    IF X > L THEN
    	DEAD_BAND := X - L;
    ELSIF X < -L THEN
    	DEAD_BAND := X + L;
    ELSE
    	DEAD_BAND := 0.0;
    END_IF

    (* revision history
    hm	2. nov. 2007	rev 1.0
    	original version

    hm	14. jun. 2008	rev 1.1
    	improved performance

    hm	18. jan. 2011	rev 1.2
    	assign 0 before return
    *)
END_FUNCTION

(* ---- DEAD_ZONE.st ---- *)
FUNCTION DEAD_ZONE
    (*http://www.oscat.de/images/OSCATBasic/oscat_basic333_en.pdf#page=394*)
    IF ABS(X) > L THEN
    	DEAD_ZONE := X;
    ELSE
    	DEAD_ZONE := 0.0;
    END_IF

    (* revision history
    hm	12. feb. 2007	rev 1.0
    	original version

    hm	14. jun. 2008	rev 1.1
    	improved performance

    hm	11. mar. 2009	rev 1.2
    	real constants updated to new systax using dot

    *)
END_FUNCTION

(* ---- DEC1.st ---- *)
FUNCTION DEC1
    (*http://www.oscat.de/images/OSCATBasic/oscat_basic333_en.pdf#page=46*)
    IF X = 0 THEN
    	DEC1 := N - 1;
    ELSE
    	DEC1 := X - 1;
    END_IF

    (* this is a very elegant version but 50% slower
    X := (X - 1 + N) MOD N;
    *)

    (* revision history
    hm	13. oct. 2008	rev 1.0
    	original version

    hm	27. oct. 2008	rev 1.1
    	added statement to return value for compatibility reasons

    *)
END_FUNCTION

(* ---- DEC_TO_BYTE.st ---- *)
FUNCTION DEC_TO_BYTE
    (*http://www.oscat.de/images/OSCATBasic/oscat_basic333_en.pdf#page=150*)
    pt ACCESS ADR(DEC);
    stop := LEN(DEC);
    FOR i := 1 TO stop DO
    	(* read the first character and subtract 48 to get value in decimal 0 = 48 *)
    	X := pt;
        intX := BYTE_TO_USINT(X);
    	(* calculate the value of the digit *)
    	IF intX > 47 AND intX < 58 THEN
    		DEC_TO_BYTE := USINT_TO_BYTE(BYTE_TO_USINT(DEC_TO_BYTE) * 10 + intX - 48);
    	END_IF
    	pt ACCESS (ADR(pt) + 1);
    END_FOR

    (* revision histroy
    hm	20. jun. 2008	rev 1.0
    	original release

    hm	30. sep.2008	rev 1.1
    	changed length of input string from 20 to 10
    	corrected an error where decoding of characters 8 and 9 would fail

    *)

END_FUNCTION

(* ---- DEC_TO_DWORD.st ---- *)
FUNCTION DEC_TO_DWORD
    (*http://www.oscat.de/images/OSCATBasic/oscat_basic333_en.pdf#page=150*)
    pt ACCESS ADR(DEC);
    stop := LEN(DEC);
    FOR i := 1 TO stop DO
    	(* read the first character and subtract 48 to get value in decimal 0 = 48 *)
    	X := pt;
        intX := BYTE_TO_USINT(X);
    	(* calculate the value of the digit *)
    	IF intX > 47 AND intX < 58 THEN
    		DEC_TO_DWORD := USINT_TO_DWORD(DWORD_TO_USINT(DEC_TO_DWORD) * 10 + intX - 48);
    	END_IF
    	pt ACCESS (ADR(pt) + 1);
    END_FOR

    (* revision histroy
    hm	20. jun. 2008	rev 1.0
    	original release

    hm	30. sep. 2008	rev 1.1
    	corrected an error where decoding of characters 8 and 9 would fail
    *)

END_FUNCTION

(* ---- DEC_TO_INT.st ---- *)
FUNCTION DEC_TO_INT
    (*http://www.oscat.de/images/OSCATBasic/oscat_basic333_en.pdf#page=151*)
    pt ACCESS ADR(DEC);
    stop := LEN(DEC);
    FOR i := 1 TO stop DO
    	(* read the first character and subtract 48 to get value in decimal 0 = 48 *)
    	X := pt;
        intX := BYTE_TO_USINT(X);
    	(* calculate the value of the digit *)
    	IF intX > 47 AND intX < 58 THEN
    		DEC_TO_INT := DEC_TO_INT * 10 + intX - 48;
    	ELSIF intX = 45 AND DEC_TO_INT = 0 THEN
    		sign := TRUE;
    	END_IF
    	pt ACCESS (ADR(pt) + 1);
    END_FOR
    IF sign THEN DEC_TO_INT := -DEC_TO_INT; END_IF

    (* revision histroy
    hm	20. jun. 2008	rev 1.0
    	original release

    hm	30. sep. 2008	rev 1.1
    	changed length of input string from 20 to 10
    	corrected an error where decoding of characters 8 and 9 would fail
    *)

END_FUNCTION

(* ---- DEG.st ---- *)
FUNCTION DEG
    (*http://www.oscat.de/images/OSCATBasic/oscat_basic333_en.pdf#page=46*)
    DEG := MODR(57.29577951308232 * RAD, 360.0);

    (* revision history
    hm	4. aug 2006	rev 1.0
    	original version

    hm 16. oct 2007	rev 1.1
    	added modr statement which prohibits DEG to become bigger than 360

    hm	10. mar. 2009	rev 1.2
    	real constants updated to new systax using dot
    *)
END_FUNCTION

(* ---- DEG_TO_DIR.st ---- *)
FUNCTION DEG_TO_DIR
    (*http://www.oscat.de/images/OSCATBasic/oscat_basic333_en.pdf#page=356*)
    IF L = 0 THEN ly := cLOCATION_DEFAULT; ELSE ly := MIN(L, cLOCATION_LMAX); END_IF
    RETVAL := cDIRS[ly, ((SHL(DEG,N-1) + 45) / 90) MOD SHL(INT#2,N)*SHR(INT#8,N)];
    DEG_TO_DIR := TRUE;

    (*
    DIR := ((SHL(DEG,N-1) + 45) / 90) MOD SHL(INT#2,N);
    explanation :
    DIR is calculated BY the following formula:
    DIR := ((DIR + 45) / 90) MOD 4 if N = 1 digit
    North = 0, East = 1 ....
    DIR := ((DIR + 22,5) / 45) MOD 8 if N = 2 digit
    convert to integer calculation
    DIR := ((DIR*2 + 45) / 90) MOD 8
    N = 0, NE = 1 ....
    ther above formula replaces 2N with shift for performance
    *)

    (* revision histroy
    hm	11. jun. 2008	rev 1.0
    	original release

    hm	22. oct. 2008	rev 1.1
    	changed size of string variables to 30
    *)
END_FUNCTION

(* ---- DEL_CHARS.st ---- *)
FUNCTION DEL_CHARS
    (*http://www.oscat.de/images/OSCATBasic/oscat_basic333_en.pdf#page=151*)
    (* copy input string *)
    RETVAL := IN;
    stop := LEN(IN);
    WHILE pos <= stop DO
    	IF FIND(CX, MID(RETVAL, 1, pos)) > 0 THEN
    		(* wrong chracter needs to be deleted *)
    		RETVAL := DELETE(RETVAL, 1, pos);
    		stop := stop - 1;	(* the string is one character shorter now *)
    	ELSE
    		(* charcter not found skip to next one *)
    		pos := pos + 1;
    	END_IF
    END_WHILE
    DEL_CHARS := TRUE;

    (* revision history

    hm		18. jun. 2008	rev 1.0
    	original version

    *)
END_FUNCTION

(* ---- DIFFER.st ---- *)
FUNCTION DIFFER
    (*http://www.oscat.de/images/OSCATBasic/oscat_basic333_en.pdf#page=47*)
    DIFFER := ABS(IN1 - IN2) > X;

    (* revision history
    hm		8. oct 2006		rev 1.0
    	original version

    hm		16. mar 2008	rev 1.1
    	improverd code for performance

    *)
END_FUNCTION

(* ---- DIR_TO_DEG.st ---- *)
FUNCTION DIR_TO_DEG
    (*http://www.oscat.de/images/OSCATBasic/oscat_basic333_en.pdf#page=360*)
    IF L = 0 THEN ly := cLOCATION_DEFAULT; ELSE ly := MIN(L, cLOCATION_LMAX); END_IF
    FOR i := 0 TO 15 DO
    	IF cDIRS[ly, i] = DIR THEN EXIT; END_IF
    END_FOR
    DIR_TO_DEG := SHR(i * 45 + 1, 1);

    (* revision histroy
    hm	22. oct. 2008	rev 1.1
    	original release

    *)
END_FUNCTION

(* ---- DST.st ---- *)
FUNCTION DST
    (*http://www.oscat.de/images/OSCATBasic/oscat_basic333_en.pdf#page=121*)
    yr := YEAR_OF_DATE(DT_TO_DATE(UTC));
    ltc := DT_TO_UDINT(UTC);
    idate := DT_TO_UDINT(SET_DT(yr, 3, 31, 1, 0, 0));
    yr4 := SHR(5 * INT_TO_UDINT(yr), 2) + 1;
    DST := (idate - ((yr4 + 3) MOD 7) * 86400 <= ltc) AND (idate + (214 - (yr4) MOD 7) * 86400 > ltc);

    (*
    Equation used TO calculate the beginning OF European Summer TIME:
    Sunday (31 - (5*y/4 + 4) mod 7) March at 01.00 UTC
    (valid through 2099, courtesy of Robert H. van Gent, EC).

    European Summer Time ends (clocks go back) at 01.00 UTC on

        * 29 October 2006
        * 28 October 2007
        * 26 October 2008

    Equation used to calculate the end of European Summer Time:
    Sunday (31 - (5*y/4 + 1) mod 7) October at 01.00 UTC
    (validity AND credits as above).

    *)

    (* revision history
    hm	4. aug 2006	rev 1.0
    	original version

    hm	24. okt 2007	rev 1.1
    	deleted time_zone_offset input because DST is generally at 01:00 UTC and not mesz
    	uk starts 01:00 UTC and also greece

    hm	1. dec 2007	rev 1.2
    	changed code to improve performance

    hm	16. mar. 2008	rev 1.3
    	added type conversion to avoid warnings under codesys 3.0
    	code improvement for better performance

    hm	7. oct. 2008	rev 1.4
    	changed name of function year to year_of_date

    hm	24. jan. 2011	rev 1.5
    	improved performance
    *)

END_FUNCTION

(* ---- DT2_TO_SDT.st ---- *)
FUNCTION DT2_TO_SDT
    (*http://www.oscat.de/images/OSCATBasic/oscat_basic333_en.pdf#page=121*)
    RETVAL.YEAR := YEAR_OF_DATE(DI);
    RETVAL.MONTH := MONTH_OF_DATE(DI);
    RETVAL.DAY := DAY_OF_MONTH(DI);
    RETVAL.WEEKDAY := DAY_OF_WEEK(DI);
    RETVAL.MS := UDINT_TO_INT(TOD_TO_UDINT(TI) MOD 1000);
    RETVAL.SECOND := UDINT_TO_INT((TOD_TO_UDINT(TI) / 1000) MOD 60);
    RETVAL.MINUTE := UDINT_TO_INT((TOD_TO_UDINT(TI) / 60000) MOD 60);
    RETVAL.HOUR := UDINT_TO_INT(TOD_TO_UDINT(TI) / 3600000);
    DT2_TO_SDT:=TRUE;
    (* revision history

    hm 18. oct. 2008	rev 1.0
    	original version

    *)
END_FUNCTION

(* ---- DT_TO_SDT.st ---- *)
FUNCTION DT_TO_SDT
    (*http://www.oscat.de/images/OSCATBasic/oscat_basic333_en.pdf#page=122*)
    tmp := DT_TO_DATE(DTI);
    tdt := DT_TO_UDINT(DTI) - DATE_TO_UDINT(tmp);
    RETVAL.YEAR := YEAR_OF_DATE(tmp);
    RETVAL.MONTH := MONTH_OF_DATE(tmp);
    RETVAL.DAY := DAY_OF_MONTH(tmp);
    RETVAL.WEEKDAY := DAY_OF_WEEK(tmp);
    RETVAL.SECOND := UDINT_TO_INT(tdt MOD 60);
    RETVAL.MINUTE := UDINT_TO_INT((tdt / 60) MOD 60);
    RETVAL.HOUR := UDINT_TO_INT(tdt / 3600);
    DT_TO_SDT:=TRUE;
    (* revision history

    hm 18. oct. 2008	rev 1.0
    	original version

    *)
END_FUNCTION

(* ---- DT_TO_STRF.st ---- *)
FUNCTION DT_TO_STRF
    (*http://www.oscat.de/images/OSCATBasic/oscat_basic333_en.pdf#page=152*)
    IF LANG < 1 THEN ly := cLANGUAGE_DEFAULT; ELSE ly := MIN(cLANGUAGE_LMAX, LANG); END_IF

    (* decode date and time information *)
    dx := DT_TO_DATE(DTI);
    td := DT_TO_TOD(DTI);

    (* parse the format string *)
    RETVAL := FMT;
    pos := FIND(RETVAL, '#');
    WHILE pos > 0 DO
    	(* retrieve format identifier *)
    	f := BYTE_TO_INT(CODE(RETVAL, pos + 1));
    	(* generate the return string according to the format character *)
    	fs := '';
    	CASE f OF
    		65 : (* letter A retunrs the year in 4 digits *)
    			fs := INT_TO_STRING(YEAR_OF_DATE(dx));
    		66 : (* letter B returns the year in exactly 2 digits *)
                fs := INT_TO_STRING(YEAR_OF_DATE(dx));
    			fs := RIGHT(fs,2);
    		67 : (* letter C returns the month with 1 or 2 digits *)
    			fs := INT_TO_STRING(MONTH_OF_DATE(dx));
    		68 : (* letter D returns the month with exactly 2 digits *)
    			fs := INT_TO_STRING(MONTH_OF_DATE(dx));
    			IF LEN(fs) < 2 THEN fs := CONCAT('0', fs); END_IF
    		69 : (* letter E returns the month with 3 characters *)
    			MONTH_TO_STRING(MONTH_OF_DATE(dx), ly, 3, fs);
    		70 : (* letter f returns the month with all characters *)
    			MONTH_TO_STRING(MONTH_OF_DATE(dx), ly, 0, fs);
    		71 : (* letter G returns the day with up to 2 digits *)
    			fs := INT_TO_STRING(DAY_OF_MONTH(dx));
    		72 : (* letter H returns the day of the month with exactly 2 digits *)
    			fs := INT_TO_STRING(DAY_OF_MONTH(dx));
    			IF LEN(fs) < 2 THEN fs := CONCAT(FILL, fs); END_IF
    		73 : (* letter I returns the weekday as the number 1..7 1 = monday *)
    			fs := INT_TO_STRING(DAY_OF_WEEK(dx));
    		74 : (* letter J returns the weekday in 2 character writing *)
    			WEEKDAY_TO_STRING(DAY_OF_WEEK(dx), ly, 2, fs);
    		75 : (* letter K returns the weekday with all characters *)
    			WEEKDAY_TO_STRING(DAY_OF_WEEK(dx), ly, 0, fs);
    		76 : (* letter L returns AM or PM for the given DateTime *)
    			IF td >= TOD#12:00 THEN fs := 'PM'; ELSE fs := 'AM'; END_IF
    		77 : (* letter M returns the hour in 1 or 2 digit form 0..24h *)
    			fs := INT_TO_STRING(HOUR(td));
    		78 : (* letter N returns the hour in exactly 2 digit form 0..24h *)
    			fs := INT_TO_STRING(HOUR(td));
    			IF LEN(fs) < 2 THEN fs := CONCAT(FILL, fs); END_IF
    		79 : (* letter O returns the hour in 1 or 2 digit form 0..12h *)
    			tmp := HOUR(td) MOD 12;
    			IF tmp = 0 THEN tmp := 12; END_IF
    			fs := INT_TO_STRING(tmp);
    		80 : (* letter P returns the hour in exactly 2 digit form 0..12h *)
    			tmp := HOUR(td) MOD 12;
    			IF tmp = 0 THEN tmp := 12; END_IF
    			fs := INT_TO_STRING(tmp);
    			IF LEN(fs) < 2 THEN fs := CONCAT(FILL, fs); END_IF
    		81 : (* letter Q returns the minute of the hour in 1 or two digit form *)
    			fs := INT_TO_STRING(MINUTE(td));
    		82 : (* letter R returns the minute of the hour in exactly two digit form *)
    			fs := INT_TO_STRING(MINUTE(td));
    			IF LEN(fs) < 2 THEN fs := CONCAT(FILL, fs); END_IF
    		83 : (* letter S returns the second of the minute in 1 or two digit form *)
    			fs := INT_TO_STRING(REAL_TO_INT(SECOND(td)));
    		84 : (* letter T returns the second of the minute in exactly two digit form *)
    			fs := INT_TO_STRING(REAL_TO_INT(SECOND(td)));
    			IF LEN(fs) < 2 THEN fs := CONCAT(FILL, fs); END_IF
    		85 : (* letter U returns the milliseconds in 1 to 3 digits *)
    			fs := INT_TO_STRING(MS);
    		86 : (* letter V returns the milliseconds in exactly 3 digit form *)
    			fs := INT_TO_STRING(MS);
    			fs := CONCAT('00',fs);
    			fs := RIGHT(fs, 3);
    		87 : (* letter W returns the day of the month with exactly 2 digits first digit is filled with BLANK if necessary *)
    			fs := INT_TO_STRING(DAY_OF_MONTH(dx));
    			IF LEN(fs) < 2 THEN fs := CONCAT(BLANK, fs); END_IF
    		88 : (* letter X returns the month with exactly 2 digits first digit is filled with BLANK if necessary *)
    			fs := INT_TO_STRING(MONTH_OF_DATE(dx));
    			IF LEN(fs) < 2 THEN fs := CONCAT(BLANK, fs); END_IF
    		END_CASE
    	RETVAL := REPLACE(RETVAL, fs, 2, pos);
    	pos := FIND(RETVAL, '#');
    END_WHILE
    DT_TO_STRF := TRUE;

    (* revision history
    hm	7. oct. 2008	rev 1.0
    	original version

    hm	19. oct. 2008	rev 1.1
    	changed language setup constants
    *)

END_FUNCTION

(* ---- DW_TO_REAL.st ---- *)
FUNCTION DW_TO_REAL
    (*http://www.oscat.de/images/OSCATBasic/oscat_basic333_en.pdf#page=225*)
    pt := ADR(X);
    DW_TO_REAL := pt;

    (* revision history
    hm	18. apr. 2008
    	original version

    *)
END_FUNCTION

(* ---- DWORD_OF_BYTE.st ---- *)
FUNCTION DWORD_OF_BYTE
    (*http://www.oscat.de/images/OSCATBasic/oscat_basic333_en.pdf#page=225*)
    DWORD_OF_BYTE := SHL(SHL(SHL(BYTE_TO_DWORD(B3),8) OR BYTE_TO_DWORD(B2),8) OR BYTE_TO_DWORD(B1),8) OR BYTE_TO_DWORD(B0);

    (* revision history
    hm	24. jan 2007	rev 1.0
    	original version

    hm 2. jan 2008	rev 1.1
    	inproved performance

    hm	23. apr. 2008	rev 1.2
    	reverse order of inputs to be more logical

    hm	18. jul. 2009	rev 1.3
    	added type conversions for compatibility reasons
    *)
END_FUNCTION

(* ---- DWORD_OF_WORD.st ---- *)
FUNCTION DWORD_OF_WORD
    (*http://www.oscat.de/images/OSCATBasic/oscat_basic333_en.pdf#page=226*)
    DWORD_OF_WORD := SHL(WORD_TO_DWORD(W1),16) OR WORD_TO_DWORD(W0);

    (* revision history

    hm	18. jul. 2009	rev 1.0
    	original version

    *)
END_FUNCTION
